{region 'Documentation'}
(*!
<summary>Selects explicit stimuli and expected results for one scenario.</summary>
*)
{endregion}
METHOD PRIVATE SelectScenario : BOOL //! TRUE after selecting a supported scenario and its literal expectations; FALSE reports an unknown scenario.
VAR
    Index : UINT;
END_VAR
SelectScenario := FALSE;
FSubjectEnable := TRUE;
FContinueScenario := FALSE;
FInput := 'A';
FExpected := 'B';
FWideInput := "A";
FWideExpected := "B";
FChar := BYTE#16#41;
FExpectedChar := BYTE#16#42;
FWideChar := WORD#16#0041;
FExpectedWideChar := WORD#16#0042;
CASE FScenario OF
    ScenarioShortQuoted:
        FExpectedMessage1 := 'Assertion failed: values are not equal. Expected = $'B$', Actual = $'A$'.';
        FExpectedMessage2 := 'Assertion failed: values are not equal. Expected = $'B$', Actual = $'A$'.';
        FExpectedMessage3 := 'Assertion failed: values are not equal. Expected = $'B$' (16#42), Actual = $'A$' (16#41).';
        FExpectedMessage4 := 'Assertion failed: values are not equal. Expected = $'B$' (16#0042), Actual = $'A$' (16#0041).';
        FTextExpectedResult := E_Result.Failed;
        FTextExpectedFinding := TRUE;
        FWideTextExpectedResult := E_Result.Failed;
        FWideTextExpectedFinding := TRUE;
        FCharacterExpectedResult := E_Result.Failed;
        FCharacterExpectedFinding := TRUE;
        FWideCharacterExpectedResult := E_Result.Failed;
        FWideCharacterExpectedFinding := TRUE;
    ScenarioPreview38:
        FInput := 'AAAAAAAAAAAAAAAAAAAAAAAAAAAAAAAAAAAAAA';
        FExpected := 'BBBBBBBBBBBBBBBBBBBBBBBBBBBBBBBBBBBBBB';
        FWideInput := "AAAAAAAAAAAAAAAAAAAAAAAAAAAAAAAAAAAAAA";
        FWideExpected := "BBBBBBBBBBBBBBBBBBBBBBBBBBBBBBBBBBBBBB";
        FExpectedMessage1 := 'Assertion failed: values are not equal. Expected = $'BBBBBBBBBBBBBBBBBBBBBBBBBBBBBBBBBBBBBB$', Actual = $'AAAAAAAAAAAAAAAAAAAAAAAAAAAAAAAAAAAAAA$'.';
        FExpectedMessage2 := 'Assertion failed: values are not equal. Expected = $'BBBBBBBBBBBBBBBBBBBBBBBBBBBBBBBBBBBBBB$', Actual = $'AAAAAAAAAAAAAAAAAAAAAAAAAAAAAAAAAAAAAA$'.';
        FExpectedMessage3 := 'Assertion failed: values are not equal. Expected = $'B$' (16#42), Actual = $'A$' (16#41).';
        FExpectedMessage4 := 'Assertion failed: values are not equal. Expected = $'B$' (16#0042), Actual = $'A$' (16#0041).';
        FTextExpectedResult := E_Result.Failed;
        FTextExpectedFinding := TRUE;
        FWideTextExpectedResult := E_Result.Failed;
        FWideTextExpectedFinding := TRUE;
        FCharacterExpectedResult := E_Result.Failed;
        FCharacterExpectedFinding := TRUE;
        FWideCharacterExpectedResult := E_Result.Failed;
        FWideCharacterExpectedFinding := TRUE;
    ScenarioPreview39:
        FInput := 'AAAAAAAAAAAAAAAAAAAAAAAAAAAAAAAAAAAAAAA';
        FExpected := 'BBBBBBBBBBBBBBBBBBBBBBBBBBBBBBBBBBBBBBB';
        FWideInput := "AAAAAAAAAAAAAAAAAAAAAAAAAAAAAAAAAAAAAAA";
        FWideExpected := "BBBBBBBBBBBBBBBBBBBBBBBBBBBBBBBBBBBBBBB";
        FExpectedMessage1 := 'Assertion failed: values are not equal. Expected = $'BBBBBBBBBBBBBBBBBBBBBBBBBBBBBBBBBBB...$', Actual = $'AAAAAAAAAAAAAAAAAAAAAAAAAAAAAAAAAAA...$'.';
        FExpectedMessage2 := 'Assertion failed: values are not equal. Expected = $'BBBBBBBBBBBBBBBBBBBBBBBBBBBBBBBBBBB...$', Actual = $'AAAAAAAAAAAAAAAAAAAAAAAAAAAAAAAAAAA...$'.';
        FExpectedMessage3 := 'Assertion failed: values are not equal. Expected = $'B$' (16#42), Actual = $'A$' (16#41).';
        FExpectedMessage4 := 'Assertion failed: values are not equal. Expected = $'B$' (16#0042), Actual = $'A$' (16#0041).';
        FTextExpectedResult := E_Result.Failed;
        FTextExpectedFinding := TRUE;
        FWideTextExpectedResult := E_Result.Failed;
        FWideTextExpectedFinding := TRUE;
        FCharacterExpectedResult := E_Result.Failed;
        FCharacterExpectedFinding := TRUE;
        FWideCharacterExpectedResult := E_Result.Failed;
        FWideCharacterExpectedFinding := TRUE;
    ScenarioDifferenceBeyondPreview:
        FInput := 'AAAAAAAAAAAAAAAAAAAAAAAAAAAAAAAAAAAAAAAX';
        FExpected := 'AAAAAAAAAAAAAAAAAAAAAAAAAAAAAAAAAAAAAAAY';
        FWideInput := "AAAAAAAAAAAAAAAAAAAAAAAAAAAAAAAAAAAAAAAX";
        FWideExpected := "AAAAAAAAAAAAAAAAAAAAAAAAAAAAAAAAAAAAAAAY";
        FExpectedMessage1 := 'Assertion failed: values are not equal. Expected = $'AAAAAAAAAAAAAAAAAAAAAAAAAAAAAAAAAAA...$', Actual = $'AAAAAAAAAAAAAAAAAAAAAAAAAAAAAAAAAAA...$'.';
        FExpectedMessage2 := 'Assertion failed: values are not equal. Expected = $'AAAAAAAAAAAAAAAAAAAAAAAAAAAAAAAAAAA...$', Actual = $'AAAAAAAAAAAAAAAAAAAAAAAAAAAAAAAAAAA...$'.';
        FExpectedMessage3 := 'Assertion failed: values are not equal. Expected = $'B$' (16#42), Actual = $'A$' (16#41).';
        FExpectedMessage4 := 'Assertion failed: values are not equal. Expected = $'B$' (16#0042), Actual = $'A$' (16#0041).';
        FTextExpectedResult := E_Result.Failed;
        FTextExpectedFinding := TRUE;
        FWideTextExpectedResult := E_Result.Failed;
        FWideTextExpectedFinding := TRUE;
        FCharacterExpectedResult := E_Result.Failed;
        FCharacterExpectedFinding := TRUE;
        FWideCharacterExpectedResult := E_Result.Failed;
        FWideCharacterExpectedFinding := TRUE;
    ScenarioAtCapacity:
        FOR Index := 0 TO Param_Assertions.AssertionStringLength - 1 DO
            // SA0175: Bounded byte writes construct exact input/terminator boundaries; no UTF-8 decoding.
            {analysis -175}
            FInput[Index] := BYTE#16#41;
            FExpected[Index] := BYTE#16#42;
            {analysis +175}
        END_FOR;
        // SA0175: Bounded byte writes construct exact input/terminator boundaries; no UTF-8 decoding.
        {analysis -175}
        FInput[Param_Assertions.AssertionStringLength] := 0;
        FExpected[Param_Assertions.AssertionStringLength] := 0;
        {analysis +175}
        FOR Index := 0 TO Param_Assertions.AssertionWStringLength - 1 DO
            FWideInput[Index] := WORD#16#0041;
            FWideExpected[Index] := WORD#16#0042;
        END_FOR;
        FWideInput[Param_Assertions.AssertionWStringLength] := 0;
        FWideExpected[Param_Assertions.AssertionWStringLength] := 0;
        FExpectedMessage1 := 'Assertion failed: values are not equal. Expected = $'BBBBBBBBBBBBBBBBBBBBBBBBBBBBBBBBBBB...$', Actual = $'AAAAAAAAAAAAAAAAAAAAAAAAAAAAAAAAAAA...$'.';
        FExpectedMessage2 := 'Assertion failed: values are not equal. Expected = $'BBBBBBBBBBBBBBBBBBBBBBBBBBBBBBBBBBB...$', Actual = $'AAAAAAAAAAAAAAAAAAAAAAAAAAAAAAAAAAA...$'.';
        FExpectedMessage3 := 'Assertion failed: values are not equal. Expected = $'B$' (16#42), Actual = $'A$' (16#41).';
        FExpectedMessage4 := 'Assertion failed: values are not equal. Expected = $'B$' (16#0042), Actual = $'A$' (16#0041).';
        FTextExpectedResult := E_Result.Failed;
        FTextExpectedFinding := TRUE;
        FWideTextExpectedResult := E_Result.Failed;
        FWideTextExpectedFinding := TRUE;
        FCharacterExpectedResult := E_Result.Failed;
        FCharacterExpectedFinding := TRUE;
        FWideCharacterExpectedResult := E_Result.Failed;
        FWideCharacterExpectedFinding := TRUE;
    ScenarioCodeFallback:
        FChar := 0;
        FExpectedChar := 1;
        FWideChar := WORD#16#0100;
        FExpectedWideChar := WORD#16#0200;
        FExpectedMessage1 := 'Assertion failed: values are not equal. Expected = $'B$', Actual = $'A$'.';
        FExpectedMessage2 := 'Assertion failed: values are not equal. Expected = $'B$', Actual = $'A$'.';
        FExpectedMessage3 := 'Assertion failed: values are not equal. Expected = 16#01, Actual = 16#00.';
        FExpectedMessage4 := 'Assertion failed: values are not equal. Expected = 16#0200, Actual = 16#0100.';
        FTextExpectedResult := E_Result.Failed;
        FTextExpectedFinding := TRUE;
        FWideTextExpectedResult := E_Result.Failed;
        FWideTextExpectedFinding := TRUE;
        FCharacterExpectedResult := E_Result.Failed;
        FCharacterExpectedFinding := TRUE;
        FWideCharacterExpectedResult := E_Result.Failed;
        FWideCharacterExpectedFinding := TRUE;
    ScenarioReplacement:
        // SA0175: Deliberately different raw bytes; both previews must render the same marker.
        {analysis -175}
        FInput := '$E4$01';
        FExpected := '$FF$7F';
        FWideInput := "$0100$20AC";
        FWideExpected := "$0001$FFFF";
        FExpectedMessage1 := 'Assertion failed: values are not equal. Expected = $'$D7$D7$', Actual = $'$D7$D7$'.';
        FExpectedMessage2 := 'Assertion failed: values are not equal. Expected = $'$D7$D7$', Actual = $'$D7$D7$'.';
        FExpectedMessage3 := 'Assertion failed: values are not equal. Expected = $'B$' (16#42), Actual = $'A$' (16#41).';
        FExpectedMessage4 := 'Assertion failed: values are not equal. Expected = $'B$' (16#0042), Actual = $'A$' (16#0041).';
        FTextExpectedResult := E_Result.Failed;
        FTextExpectedFinding := TRUE;
        FWideTextExpectedResult := E_Result.Failed;
        FWideTextExpectedFinding := TRUE;
        FCharacterExpectedResult := E_Result.Failed;
        FCharacterExpectedFinding := TRUE;
        FWideCharacterExpectedResult := E_Result.Failed;
        FWideCharacterExpectedFinding := TRUE;
        {analysis +175}
ELSE
    Error(Message := 'Unknown Assertion scenario.');
    RETURN;
END_CASE;
SelectScenario := TRUE;
END_METHOD

END_FUNCTION_BLOCK

// ---- Framework/Assertions/POU/Utilities/CreateAssertionTextValue_String.TcPOU
{region 'Documentation'}
(*!
<summary>Render a quoted diagnostic preview with at most AssertionValueLength output bytes.
Printable ASCII is retained; other code units become byte 16#D7 without expansion.</summary>
<description>
Zero terminates the input. Quotes and backslashes remain literal. Shortening reserves
space for enclosing quotes and an ellipsis; the default limit retains 35 code units.
Rendering is lossy and does not alter the compared input or its result.
</description>
*)
{endregion}
FUNCTION INTERNAL CreateAssertionTextValue_String : STRING(GVL_Constants.AssertionValueLength) //! Bounded diagnostic aid; not a lossless representation for subsequent comparison.
VAR_INPUT
    Value : STRING(GVL_Constants.MessageLength); //! Text to preview; zero terminates the input.
END_VAR
VAR
    Text : STRING(GVL_Constants.AssertionValueLength);
    CharacterIndex : INT;
    CopyLength : INT;
    Code : BYTE;
    Shortened : BOOL;
END_VAR
VAR CONSTANT
    Quote : STRING(1) := '$'';
    Ellipsis : STRING(3) := '...';
    QuoteLength : INT := 2;
    EllipsisLength : INT := 3;
    FirstPrintableAscii : BYTE := 16#20;
    LastPrintableAscii : BYTE := 16#7E;
    ReplacementByte : BYTE := 16#D7;
END_VAR

CopyLength := UINT_TO_INT(GVL_Constants.AssertionValueLength) - QuoteLength;
// SA0175: Bounded diagnostic code-unit rendering; each unsupported unit becomes one byte.
{analysis -175}
Shortened := TRUE;
FOR CharacterIndex := 0 TO CopyLength DO
    IF Value[CharacterIndex] = 0 THEN
        CopyLength := CharacterIndex;
        Shortened := FALSE;
        EXIT;
    END_IF;
END_FOR;
IF Shortened THEN
    CopyLength := CopyLength - EllipsisLength;
END_IF;

FOR CharacterIndex := 0 TO CopyLength - 1 DO
    Code := Value[CharacterIndex];
    IF (Code >= FirstPrintableAscii) AND (Code <= LastPrintableAscii) THEN
        Text[CharacterIndex] := Code;
    ELSE
        Text[CharacterIndex] := ReplacementByte;
    END_IF;
END_FOR;
Text[CopyLength] := 0;
{analysis +175}

IF Shortened THEN
    Text := CONCAT(Text, Ellipsis);
END_IF;
CreateAssertionTextValue_String := CONCAT(Quote, Text);
CreateAssertionTextValue_String := CONCAT(CreateAssertionTextValue_String, Quote);

END_FUNCTION

// ---- Framework/Assertions/POU/Utilities/CreateAssertionTextValue_WString.TcPOU
{region 'Documentation'}
(*!
<summary>Render a quoted diagnostic preview with at most AssertionValueLength output bytes.
Printable ASCII is retained; other code units become byte 16#D7 without expansion.</summary>
<description>
Zero terminates the input. Quotes and backslashes remain literal. Shortening reserves
space for enclosing quotes and an ellipsis; the default limit retains 35 code units.
Rendering is lossy and does not alter the compared input or its result.
</description>
*)
{endregion}
FUNCTION INTERNAL CreateAssertionTextValue_WString : STRING(GVL_Constants.AssertionValueLength) //! Bounded diagnostic aid; not a lossless representation for subsequent comparison.
VAR_INPUT
    Value : WSTRING(GVL_Constants.MessageLength); //! Text to preview; zero terminates the input.
END_VAR
VAR
    Text : STRING(GVL_Constants.AssertionValueLength);
    CharacterIndex : INT;
    CopyLength : INT;
    Code : WORD;
    Shortened : BOOL;
END_VAR
VAR CONSTANT
    Quote : STRING(1) := '$'';
    Ellipsis : STRING(3) := '...';
    QuoteLength : INT := 2;
    EllipsisLength : INT := 3;
    FirstPrintableAscii : WORD := 16#20;
    LastPrintableAscii : WORD := 16#7E;
    ReplacementByte : BYTE := 16#D7;
END_VAR

CopyLength := UINT_TO_INT(GVL_Constants.AssertionValueLength) - QuoteLength;
// SA0175: Bounded diagnostic code-unit rendering; each unsupported unit becomes one byte.
{analysis -175}
Shortened := TRUE;
FOR CharacterIndex := 0 TO CopyLength DO
    IF Value[CharacterIndex] = 0 THEN
        CopyLength := CharacterIndex;
        Shortened := FALSE;
        EXIT;
    END_IF;
END_FOR;
IF Shortened THEN
    CopyLength := CopyLength - EllipsisLength;
END_IF;

FOR CharacterIndex := 0 TO CopyLength - 1 DO
    Code := Value[CharacterIndex];
    IF (Code >= FirstPrintableAscii) AND (Code <= LastPrintableAscii) THEN
        Text[CharacterIndex] := WORD_TO_BYTE(Code);
    ELSE
        Text[CharacterIndex] := ReplacementByte;
    END_IF;
END_FOR;
Text[CopyLength] := 0;
{analysis +175}

IF Shortened THEN
    Text := CONCAT(Text, Ellipsis);
END_IF;
CreateAssertionTextValue_WString := CONCAT(Quote, Text);
CreateAssertionTextValue_WString := CONCAT(CreateAssertionTextValue_WString, Quote);

END_FUNCTION

// ---- Framework/Assertions/POU/Utilities/CreateAssertionTextValue_ByteArray.TcPOU
{region 'Documentation'}
(*!
<summary>Render a quoted printable-ASCII/16#D7 preview of an array range without modifying its storage. Invalid or empty ranges return two quotes. Zero and other unsupported elements become one replacement byte each. Work is bounded by the preview capacity.</summary>
*)
{endregion}
FUNCTION INTERNAL CreateAssertionTextValue_ByteArray : STRING(GVL_Constants.AssertionValueLength) //! Bounded diagnostic text; not a value for subsequent numeric comparison.
VAR_INPUT
    StartIndex : DINT; //! First selected index in Value, using the array's declared index range.
    Length : UINT; //! Number of selected elements starting at StartIndex; must fit the array range.
END_VAR
VAR_IN_OUT CONSTANT
    Value : ARRAY[*] OF BYTE; //! Read-only source array; StartIndex and Length select the diagnostic preview.
END_VAR
VAR
    LowerIndex : DINT;
    UpperIndex : DINT;
    CopyLength : INT;
    Offset : INT;
    Code : BYTE;
    Text : STRING(GVL_Constants.AssertionValueLength);
    Preview : STRING(GVL_Constants.AssertionValueLength);
END_VAR
VAR CONSTANT
    Quote : STRING(1) := '$'';
    Ellipsis : STRING(3) := '...';
    QuoteLength : INT := 2;
    EllipsisLength : INT := 3;
    FirstPrintableAscii : BYTE := 16#20;
    LastPrintableAscii : BYTE := 16#7E;
    ReplacementByte : BYTE := 16#D7;
END_VAR

CreateAssertionTextValue_ByteArray := CONCAT(Quote, Quote);
LowerIndex := LOWER_BOUND(Value, 1);
UpperIndex := UPPER_BOUND(Value, 1);

IF Length = 0 OR StartIndex < LowerIndex OR StartIndex > UpperIndex THEN
    RETURN;
END_IF;

IF UINT_TO_LINT(Length) > DINT_TO_LINT(UpperIndex) - DINT_TO_LINT(StartIndex) + 1 THEN
    RETURN;
END_IF;

IF Length > GVL_Constants.AssertionValueLength - INT_TO_UINT(QuoteLength) THEN
    CopyLength := UINT_TO_INT(GVL_Constants.AssertionValueLength) - QuoteLength - EllipsisLength;
ELSE
    CopyLength := UINT_TO_INT(Length);
END_IF;

// SA0175: Range guards bound reads; preview writes fit capacity, including the terminator.
{analysis -175}
FOR Offset := 0 TO CopyLength - 1 DO
    Code := Value[StartIndex + INT_TO_DINT(Offset)];
    IF (Code >= FirstPrintableAscii) AND (Code <= LastPrintableAscii) THEN
        Text[Offset] := Code;
    ELSE
        Text[Offset] := ReplacementByte;
    END_IF;
END_FOR;
Text[CopyLength] := 0;
{analysis +175}

Preview := Text;
IF Length > GVL_Constants.AssertionValueLength - INT_TO_UINT(QuoteLength) THEN
    Preview := CONCAT(Preview, Ellipsis);
END_IF;

CreateAssertionTextValue_ByteArray := CONCAT(Quote, Preview);
CreateAssertionTextValue_ByteArray := CONCAT(CreateAssertionTextValue_ByteArray, Quote);

END_FUNCTION

// ---- Framework/Assertions/POU/Utilities/CreateAssertionTextValue_WordArray.TcPOU
{region 'Documentation'}
(*!
<summary>Render a quoted printable-ASCII/16#D7 preview of an array range without modifying its storage. Invalid or empty ranges return two quotes. Zero and other unsupported elements become one replacement byte each. Work is bounded by the preview capacity.</summary>
*)
{endregion}
FUNCTION INTERNAL CreateAssertionTextValue_WordArray : STRING(GVL_Constants.AssertionValueLength) //! Bounded diagnostic text; not a value for subsequent numeric comparison.
VAR_INPUT
    StartIndex : DINT; //! First selected index in Value, using the array's declared index range.
    Length : UINT; //! Number of selected elements starting at StartIndex; must fit the array range.
END_VAR
VAR_IN_OUT CONSTANT
    Value : ARRAY[*] OF WORD; //! Read-only source array; StartIndex and Length select the diagnostic preview.
END_VAR
VAR
    LowerIndex : DINT;
    UpperIndex : DINT;
    CopyLength : INT;
    Offset : INT;
    Code : WORD;
    Text : STRING(GVL_Constants.AssertionValueLength);
    Preview : STRING(GVL_Constants.AssertionValueLength);
END_VAR
VAR CONSTANT
    Quote : STRING(1) := '$'';
    Ellipsis : STRING(3) := '...';
    QuoteLength : INT := 2;
    EllipsisLength : INT := 3;
    FirstPrintableAscii : WORD := 16#20;
    LastPrintableAscii : WORD := 16#7E;
    ReplacementByte : BYTE := 16#D7;
END_VAR

CreateAssertionTextValue_WordArray := CONCAT(Quote, Quote);
LowerIndex := LOWER_BOUND(Value, 1);
UpperIndex := UPPER_BOUND(Value, 1);

IF Length = 0 OR StartIndex < LowerIndex OR StartIndex > UpperIndex THEN
    RETURN;
END_IF;

IF UINT_TO_LINT(Length) > DINT_TO_LINT(UpperIndex) - DINT_TO_LINT(StartIndex) + 1 THEN
    RETURN;
END_IF;

IF Length > GVL_Constants.AssertionValueLength - INT_TO_UINT(QuoteLength) THEN
    CopyLength := UINT_TO_INT(GVL_Constants.AssertionValueLength) - QuoteLength - EllipsisLength;
ELSE
    CopyLength := UINT_TO_INT(Length);
END_IF;

// SA0175: Range guards bound reads; preview writes fit capacity, including the terminator.
{analysis -175}
FOR Offset := 0 TO CopyLength - 1 DO
    Code := Value[StartIndex + INT_TO_DINT(Offset)];
    IF (Code >= FirstPrintableAscii) AND (Code <= LastPrintableAscii) THEN
        Text[Offset] := WORD_TO_BYTE(Code);
    ELSE
        Text[Offset] := ReplacementByte;
    END_IF;
END_FOR;
Text[CopyLength] := 0;
{analysis +175}

Preview := Text;
IF Length > GVL_Constants.AssertionValueLength - INT_TO_UINT(QuoteLength) THEN
    Preview := CONCAT(Preview, Ellipsis);
END_IF;

CreateAssertionTextValue_WordArray := CONCAT(Quote, Preview);
CreateAssertionTextValue_WordArray := CONCAT(CreateAssertionTextValue_WordArray, Quote);

END_FUNCTION

// ---- Framework/Assertions/POU/Utilities/CreateAssertionTextValue_WChar.TcPOU
{region 'Documentation'}
(*!
<summary>Formats printable ASCII as a quoted character and hexadecimal code; other values as code only. Output is ASCII and at most 13 characters.</summary>
*)
{endregion}
FUNCTION INTERNAL CreateAssertionTextValue_WChar : STRING(13) //! Bounded diagnostic text; not a value for subsequent numeric comparison.
VAR_INPUT
    Value : WORD; //! Character code to render; no character validation is performed.
END_VAR
VAR
    HexText : STRING(7);
    Text : STRING(13);
END_VAR
VAR CONSTANT
    FirstPrintableAscii : WORD := 16#20;
    LastPrintableAscii : WORD := 16#7E;
    HexDigitCount : USINT := 4;
END_VAR

HexText := CreateAssertionTextValue_Hex(Value := WORD_TO_LWORD(Value),
    DigitCount := HexDigitCount);

IF (Value < FirstPrintableAscii) OR (Value > LastPrintableAscii) THEN
    CreateAssertionTextValue_WChar := HexText;
    RETURN;
END_IF;

Text := '$' $' (';
// SA0175: Printable-ASCII guard; index 1 fits the quoted template.
{analysis -175}
Text[1] := WORD_TO_BYTE(Value);
{analysis +175}
Text := CONCAT(Text, HexText);
CreateAssertionTextValue_WChar := CONCAT(Text, ')');

END_FUNCTION

// ---- SelfTests/TestCases/TestSuite_AssertionText/Test_AssertionValueTokenCount.TcPOU
{region 'Documentation'}
(*!
<summary>Checks masked BYTE/WORD token counts, count predicates and retained observations.</summary>
<description>
Literal counts distinguish full masks, selected bits, zero mask and sliced ranges.
Dedicated continuation scenarios check disabled/Failed count retention and clearing
on invalid range. Every independent scenario verifies count clearing on Reset.
Independent scenarios occupy two calls: bound Reset, then evaluation.
ProcessAssertions checks each call before ProcessTests advances. Literal expected
results belong to SelectScenario, not to a copy of the production comparison.
The local capture is cleared before each call and checked in subject-call order.
FirstFailedScenario and FailedDuringEvaluation retain the first mismatch.
Continuation scenarios explicitly retain the prior subject state. The Test Case
owns all input storage; no invalid or dangling references are constructed.
</description>
*)
{endregion}
FUNCTION_BLOCK Test_AssertionValueTokenCount EXTENDS TestCaseBase
VAR
    FEqual : AssertValueTokenCntEqual_Byte;
    FEqualExpectedResult : E_Result;
    FWideEqual : AssertValueTokenCntEqual_Word;
    FWideEqualExpectedResult : E_Result;
    FNone : AssertNoValueToken_Byte;
    FNoneExpectedResult : E_Result;
    FWideRange : AssertValueTokenCntInRange_Word;
    FWideRangeExpectedResult : E_Result;
    FData : ARRAY[-2..3] OF BYTE;
    FDataBefore : ARRAY[-2..3] OF BYTE;
    FWideData : ARRAY[-2..3] OF WORD;
    FWideDataBefore : ARRAY[-2..3] OF WORD;
    FStartIndex : DINT;
    FLength : USINT;
    FExpected : UINT;
    FMinimum : UINT;
    FMaximum : UINT;
    FToken : BYTE;
    FWideToken : WORD;
    FMask : BYTE;
    FWideMask : WORD;
    FSubjectEnable : BOOL;
    FContinueScenario : BOOL;
    FEqualExpectedFinding : BOOL;
    FEqualExpectedCount : UINT;
    FWideEqualExpectedFinding : BOOL;
    FWideEqualExpectedCount : UINT;
    FNoneExpectedFinding : BOOL;
    FNoneExpectedCount : UINT;
    FWideRangeExpectedFinding : BOOL;
    FWideRangeExpectedCount : UINT;
    FCapture : EventBuffer;
    FEvents : ARRAY[1..CaptureLength] OF ST_Event;
    FCaptureFifo : ST_FifoStatus;
    FCaptureStatus : ST_EventBufferStatus;
    FSetupValid : BOOL;
    FScenario : UINT;
    FChecked : BOOL;
    FEvaluateSubjects : BOOL;
    FObservationReady : BOOL;
    FFirstFailedScenario : UINT;
    FFailedDuringEvaluation : BOOL;
    FResultsMatch : BOOL;
    FResults : AssertTrue;
    FActivityMatch : BOOL;
    FActivity : AssertTrue;
    FInputsMatch : BOOL;
    FInputs : AssertTrue;
    FFindingsMatch : BOOL;
    FFindings : AssertTrue;
END_VAR
VAR CONSTANT
    CaptureLength : UINT := 8;
    ScenarioExactCount : UINT := 1;
    ScenarioMasked : UINT := 2;
    ScenarioZeroMask : UINT := 3;
    ScenarioSelectedBounds : UINT := 4;
    ScenarioLastElement : UINT := 5;
    ScenarioAbsent : UINT := 6;
    ScenarioFailedCount : UINT := 7;
    ScenarioDisabledRetention : UINT := 8;
    ScenarioFailedRetention : UINT := 9;
    ScenarioErrorClearsCount : UINT := 10;
    ScenarioResetAfterError : UINT := 11;
    ScenarioBelowArray : UINT := 12;
    ScenarioEndOutsideArray : UINT := 13;
    ScenarioReversedCountBounds : UINT := 14;
    LastScenario : UINT := ScenarioReversedCountBounds;
END_VAR

SUPER^();

{region 'Documentation'}
(*!
<summary>Aggregates only outer checks, not intentionally failing subjects.</summary>
*)
{endregion}
METHOD PROTECTED AggregateResults
VAR_INPUT
    Aggregator : I_ResultAggregator; //! Borrowed result sink owned by the outer Test Case; add this test's checking Assertions without resetting or retaining the sink.
END_VAR
Aggregator.AddProvider(Provider := FResults);
Aggregator.AddProvider(Provider := FActivity);
Aggregator.AddProvider(Provider := FInputs);
Aggregator.AddProvider(Provider := FFindings);
END_METHOD

{region 'Documentation'}
(*!
<summary>Calls each inherited production subject once with caller-owned input storage.</summary>
*)
{endregion}
METHOD PRIVATE CallSubjects
FEqual(Enable := FSubjectEnable,
    State := E_State.Running,
    StartIndex := FStartIndex,
    Length := FLength,
    Expected := FExpected,
    Token := FToken,
    Mask := FMask,
    IN := FData);
FWideEqual(Enable := FSubjectEnable,
    State := E_State.Running,
    StartIndex := FStartIndex,
    Length := FLength,
    Expected := FExpected,
    Token := FWideToken,
    Mask := FWideMask,
    IN := FWideData);
FNone(Enable := FSubjectEnable,
    State := E_State.Running,
    StartIndex := FStartIndex,
    Length := FLength,
    Token := FToken,
    Mask := FMask,
    IN := FData);
FWideRange(Enable := FSubjectEnable,
    State := E_State.Running,
    StartIndex := FStartIndex,
    Length := FLength,
    Minimum := FMinimum,
    Maximum := FMaximum,
    Token := FWideToken,
    Mask := FWideMask,
    IN := FWideData);
END_METHOD

{region 'Documentation'}
(*!
<summary>Checks one subject finding in call order; expected outcomes come from the scenario.</summary>
*)
{endregion}
METHOD PRIVATE CheckFinding : BOOL //! TRUE when the required finding checks pass; calls requiring no finding also succeed.
VAR_INPUT
    Subject : I_Assertion; //! Assertion interface supplying the expected finding identity.
    ExpectedResult : E_Result; //! Independently authored result expected in the captured finding.
    ExpectedFinding : BOOL; //! TRUE when this scenario requires a finding during active evaluation.
END_VAR
VAR_IN_OUT
    Index : UINT; //! One-based next finding index; advanced when this call checks a required finding.
END_VAR
CheckFinding := TRUE;
IF FEvaluateSubjects AND ExpectedFinding THEN
    CheckFinding := (FEvents[Index].SequenceId = UINT_TO_UDINT(Index))
        AND (FEvents[Index].Name = Subject.Name)
        AND (FEvents[Index].OwnerScope = E_OwnerScope.Assertion)
        AND (FEvents[Index].EventType = E_EventType.Result)
        AND (FEvents[Index].State = E_State.Running)
        AND (FEvents[Index].Result = ExpectedResult)
        AND (FEvents[Index].Message <> '');
    Index := Index + 1;
END_IF;
END_METHOD

{region 'Documentation'}
(*!
<summary>Checks exact finding count and identities; at most one finding per subject.</summary>
*)
{endregion}
METHOD PRIVATE CheckFindings
VAR
    Index : UINT;
    Matches : BOOL;
END_VAR
Index := 1;
FFindingsMatch := TRUE;
Matches := CheckFinding(Subject := FEqual,
    ExpectedResult := FEqualExpectedResult,
    ExpectedFinding := FEqualExpectedFinding,
    Index := Index);
FFindingsMatch := FFindingsMatch AND Matches;
Matches := CheckFinding(Subject := FWideEqual,
    ExpectedResult := FWideEqualExpectedResult,
    ExpectedFinding := FWideEqualExpectedFinding,
    Index := Index);
FFindingsMatch := FFindingsMatch AND Matches;
Matches := CheckFinding(Subject := FNone,
    ExpectedResult := FNoneExpectedResult,
    ExpectedFinding := FNoneExpectedFinding,
    Index := Index);
FFindingsMatch := FFindingsMatch AND Matches;
Matches := CheckFinding(Subject := FWideRange,
    ExpectedResult := FWideRangeExpectedResult,
    ExpectedFinding := FWideRangeExpectedFinding,
    Index := Index);
FFindingsMatch := FFindingsMatch AND Matches;
FFindingsMatch := FFindingsMatch
    AND (FCaptureStatus.SequenceId = UINT_TO_UDINT(Index - 1))
    AND (FCaptureStatus.LostEventCount = 0);
IF FEvaluateSubjects AND (FScenario = ScenarioFailedCount) THEN
    // SA0175: Fixed byte-substring checks of bounded diagnostic messages; no character offsets.
    {analysis -175}
    FFindingsMatch := FFindingsMatch
        AND (FIND(FEvents[1].Message, 'Actual = 2') > 0)
        AND (FIND(FEvents[4].Message, 'Actual = 2') > 0);
    {analysis +175}
END_IF;
END_METHOD

{region 'Documentation'}
(*!
<summary>Rejects incomplete subject, capture or outer Assertion setup.</summary>
*)
{endregion}
METHOD PROTECTED CheckInitialization : BOOL //! TRUE when the inherited initialization check and this concrete fixture check both accept the setup.
CheckInitialization := SUPER^.CheckInitialization();
IF NOT CheckInitialization THEN
    RETURN;
END_IF;

CheckInitialization := FSetupValid
    AND FResults.IsInitialized
    AND FActivity.IsInitialized
    AND FInputs.IsInitialized
    AND FFindings.IsInitialized;
IF NOT CheckInitialization THEN
    EventPublisher.PublishEvent(Event := CreateFrameworkEvent(Name := Name,
        ResourceName := '',
        State := State,
        Severity := E_EventSeverity.Error,
        Message := 'Text selftest setup failed.'));
END_IF;
END_METHOD

{region 'Documentation'}
(*!
<summary>Checks literal evaluation results, or NotEvaluated on the reset call.</summary>
*)
{endregion}
METHOD PRIVATE CheckResults
IF FEvaluateSubjects THEN
    FResultsMatch := (FEqual.Result = FEqualExpectedResult)
        AND (FWideEqual.Result = FWideEqualExpectedResult)
        AND (FNone.Result = FNoneExpectedResult)
        AND (FWideRange.Result = FWideRangeExpectedResult);
ELSE
    FResultsMatch := (FEqual.Result = E_Result.NotEvaluated)
        AND (FWideEqual.Result = E_Result.NotEvaluated)
        AND (FNone.Result = E_Result.NotEvaluated)
        AND (FWideRange.Result = E_Result.NotEvaluated);
END_IF;
FActivityMatch := (FEqual.Enabled = FSubjectEnable)
    AND (FEqual.ObservationActive = (FEvaluateSubjects AND FSubjectEnable))
    AND (FEqual.EvaluationActive = (FEvaluateSubjects AND FSubjectEnable))
    AND (FWideEqual.Enabled = FSubjectEnable)
    AND (FWideEqual.ObservationActive = (FEvaluateSubjects AND FSubjectEnable))
    AND (FWideEqual.EvaluationActive = (FEvaluateSubjects AND FSubjectEnable))
    AND (FNone.Enabled = FSubjectEnable)
    AND (FNone.ObservationActive = (FEvaluateSubjects AND FSubjectEnable))
    AND (FNone.EvaluationActive = (FEvaluateSubjects AND FSubjectEnable))
    AND (FWideRange.Enabled = FSubjectEnable)
    AND (FWideRange.ObservationActive = (FEvaluateSubjects AND FSubjectEnable))
    AND (FWideRange.EvaluationActive = (FEvaluateSubjects AND FSubjectEnable));
IF FEvaluateSubjects THEN
    FResultsMatch := FResultsMatch
        AND (FEqual.TokenCount = FEqualExpectedCount)
        AND (FWideEqual.TokenCount = FWideEqualExpectedCount)
        AND (FNone.TokenCount = FNoneExpectedCount)
        AND (FWideRange.TokenCount = FWideRangeExpectedCount);
ELSE
    FResultsMatch := FResultsMatch
        AND (FEqual.TokenCount = 0)
        AND (FWideEqual.TokenCount = 0)
        AND (FNone.TokenCount = 0)
        AND (FWideRange.TokenCount = 0);
END_IF;
END_METHOD

{region 'Documentation'}
(*!
<summary>Initializes outer checks and isolates intentional subject findings.</summary>
*)
{endregion}
METHOD PROTECTED Configure
VAR
    Initialized : BOOL;
END_VAR
FPreparationStateCount := 0;
FTestStateCount := 1;
FResults.Initialize(Parent := THIS^,
    AssertionName := 'Results');
FActivity.Initialize(Parent := THIS^,
    AssertionName := 'Activity');
FInputs.Initialize(Parent := THIS^,
    AssertionName := 'Inputs');
FFindings.Initialize(Parent := THIS^,
    AssertionName := 'Findings');
FSetupValid := FCapture.Initialize(Buffer := FEvents,
    FifoControl := FCaptureFifo,
    Status := FCaptureStatus);
FEqual.BindPublisher(Publisher := FCapture);
Initialized := FEqual.Initialize(Parent := THIS^,
    AssertionName := 'Equal');
FSetupValid := FSetupValid AND Initialized;
FWideEqual.BindPublisher(Publisher := FCapture);
Initialized := FWideEqual.Initialize(Parent := THIS^,
    AssertionName := 'WideEqual');
FSetupValid := FSetupValid AND Initialized;
FNone.BindPublisher(Publisher := FCapture);
Initialized := FNone.Initialize(Parent := THIS^,
    AssertionName := 'None');
FSetupValid := FSetupValid AND Initialized;
FWideRange.BindPublisher(Publisher := FCapture);
Initialized := FWideRange.Initialize(Parent := THIS^,
    AssertionName := 'WideRange');
FSetupValid := FSetupValid AND Initialized;
END_METHOD

{region 'Documentation'}
(*!
<summary>Completes abort; no asynchronous resource is owned.</summary>
*)
{endregion}
METHOD PROTECTED ProcessAbort
VAR_INPUT
    Enable : BOOL; //! Phase permission supplied by the owning Test Case; FALSE does not authorize progression, while observation may continue.
END_VAR
IF Enable THEN
    CompleteAbort();
END_IF;
END_METHOD

{region 'Documentation'}
(*!
<summary>Latches this call's checks before progression is permitted.</summary>
*)
{endregion}
METHOD PROTECTED ProcessAssertions
VAR_INPUT
    Enable : BOOL; //! Phase permission supplied by the owning Test Case; FALSE does not authorize progression, while observation may continue.
END_VAR
VAR
    Check : BOOL;
END_VAR
Check := Enable AND FObservationReady;
FResults(Enable := Check,
    State := State,
    IN := FResultsMatch);
FActivity(Enable := Check,
    State := State,
    IN := FActivityMatch);
FInputs(Enable := Check,
    State := State,
    IN := FInputsMatch);
FFindings(Enable := Check,
    State := State,
    IN := FFindingsMatch);
IF Check THEN
    FChecked := TRUE;
END_IF;
END_METHOD

{region 'Documentation'}
(*!
<summary>No Preparation phase is needed.</summary>
*)
{endregion}
METHOD PROTECTED ProcessPreparations
VAR_INPUT
    // SA0033: Required hook; this test has no Preparation phase.
    {attribute 'analysis' := '-33'}
    Enable : BOOL; //! Phase permission supplied by the owning Test Case; FALSE does not authorize progression, while observation may continue.
END_VAR
END_METHOD

{region 'Documentation'}
(*!
<summary>Restarts the scenario sequence and outer checks.</summary>
*)
{endregion}
METHOD PROTECTED ProcessReset
FScenario := ScenarioExactCount;
FChecked := FALSE;
FSubjectEnable := FALSE;
FContinueScenario := FALSE;
FEvaluateSubjects := FALSE;
FObservationReady := FALSE;
FFirstFailedScenario := 0;
FFailedDuringEvaluation := FALSE;
FCapture.Reset();
ResetSubjects();
FResults.Reset();
FActivity.Reset();
FInputs.Reset();
FFindings.Reset();
CompleteReset();
END_METHOD

{region 'Documentation'}
(*!
<summary>Consumes reset before each independent scenario; continuation retains subject state.</summary>
*)
{endregion}
METHOD PROTECTED ProcessTests
VAR_INPUT
    Enable : BOOL; //! Phase permission supplied by the owning Test Case; FALSE does not authorize progression, while observation may continue.
END_VAR
IF NOT Enable THEN
    RETURN;
END_IF;

IF FChecked THEN
    FChecked := FALSE;
    FObservationReady := FALSE;
    IF FEvaluateSubjects THEN
        IF FScenario = LastScenario THEN
            CompleteTests();
            RETURN;
        END_IF;
        FScenario := FScenario + 1;
    END_IF;
    FEvaluateSubjects := NOT FEvaluateSubjects;
END_IF;

IF NOT SelectScenario() THEN
    RETURN;
END_IF;
IF FContinueScenario THEN
    FEvaluateSubjects := TRUE;
END_IF;
FCapture.Reset();
IF NOT FEvaluateSubjects THEN
    ResetSubjects();
END_IF;
FDataBefore := FData;
FWideDataBefore := FWideData;
CallSubjects();
CheckResults();
FInputsMatch := (FData[-2] = FDataBefore[-2])
    AND (FData[-1] = FDataBefore[-1])
    AND (FData[0] = FDataBefore[0])
    AND (FData[1] = FDataBefore[1])
    AND (FData[2] = FDataBefore[2])
    AND (FData[3] = FDataBefore[3])
    AND (FWideData[-2] = FWideDataBefore[-2])
    AND (FWideData[-1] = FWideDataBefore[-1])
    AND (FWideData[0] = FWideDataBefore[0])
    AND (FWideData[1] = FWideDataBefore[1])
    AND (FWideData[2] = FWideDataBefore[2])
    AND (FWideData[3] = FWideDataBefore[3]);
CheckFindings();
IF (FFirstFailedScenario = 0)
    AND NOT (FResultsMatch AND FActivityMatch AND FInputsMatch AND FFindingsMatch) THEN
    FFirstFailedScenario := FScenario;
    FFailedDuringEvaluation := FEvaluateSubjects;
END_IF;
FObservationReady := TRUE;
END_METHOD

{region 'Documentation'}
(*!
<summary>Queues reset; the next bound FB call consumes it without evaluating.</summary>
*)
{endregion}
METHOD PRIVATE ResetSubjects
FEqual.Reset();
FWideEqual.Reset();
FNone.Reset();
FWideRange.Reset();
END_METHOD

{region 'Documentation'}
(*!
<summary>Selects explicit stimuli and expected results for one scenario.</summary>
*)
{endregion}
METHOD PRIVATE SelectScenario : BOOL //! TRUE after selecting a supported scenario and its literal expectations; FALSE reports an unknown scenario.
SelectScenario := FALSE;
FSubjectEnable := TRUE;
FContinueScenario := FALSE;
FData[-2] := BYTE#16#10;
FData[-1] := BYTE#16#21;
FData[0] := BYTE#16#11;
FData[1] := BYTE#16#20;
FData[2] := BYTE#16#11;
FData[3] := BYTE#16#99;
FWideData[-2] := WORD#16#0110;
FWideData[-1] := WORD#16#0121;
FWideData[0] := WORD#16#0111;
FWideData[1] := WORD#16#0220;
FWideData[2] := WORD#16#0111;
FWideData[3] := WORD#16#0099;
FStartIndex := -2;
FLength := 6;
FExpected := 2;
FMinimum := 2;
FMaximum := 2;
FToken := BYTE#16#11;
FWideToken := WORD#16#0111;
FMask := BYTE#16#FF;
FWideMask := WORD#16#FFFF;
CASE FScenario OF
    ScenarioExactCount:
        FEqualExpectedResult := E_Result.Passed;
        FEqualExpectedFinding := FALSE;
        FEqualExpectedCount := 2;
        FWideEqualExpectedResult := E_Result.Passed;
        FWideEqualExpectedFinding := FALSE;
        FWideEqualExpectedCount := 2;
        FNoneExpectedResult := E_Result.Failed;
        FNoneExpectedFinding := TRUE;
        FNoneExpectedCount := 2;
        FWideRangeExpectedResult := E_Result.Passed;
        FWideRangeExpectedFinding := FALSE;
        FWideRangeExpectedCount := 2;
    ScenarioMasked:
        FMask := BYTE#16#0F;
        FWideMask := WORD#16#000F;
        FExpected := 3;
        FMinimum := 3;
        FMaximum := 3;
        FEqualExpectedResult := E_Result.Passed;
        FEqualExpectedFinding := FALSE;
        FEqualExpectedCount := 3;
        FWideEqualExpectedResult := E_Result.Passed;
        FWideEqualExpectedFinding := FALSE;
        FWideEqualExpectedCount := 3;
        FNoneExpectedResult := E_Result.Failed;
        FNoneExpectedFinding := TRUE;
        FNoneExpectedCount := 3;
        FWideRangeExpectedResult := E_Result.Passed;
        FWideRangeExpectedFinding := FALSE;
        FWideRangeExpectedCount := 3;
    ScenarioZeroMask:
        FMask := 0;
        FWideMask := 0;
        FExpected := 6;
        FMinimum := 6;
        FMaximum := 6;
        FEqualExpectedResult := E_Result.Passed;
        FEqualExpectedFinding := FALSE;
        FEqualExpectedCount := 6;
        FWideEqualExpectedResult := E_Result.Passed;
        FWideEqualExpectedFinding := FALSE;
        FWideEqualExpectedCount := 6;
        FNoneExpectedResult := E_Result.Failed;
        FNoneExpectedFinding := TRUE;
        FNoneExpectedCount := 6;
        FWideRangeExpectedResult := E_Result.Passed;
        FWideRangeExpectedFinding := FALSE;
        FWideRangeExpectedCount := 6;
    ScenarioSelectedBounds:
        FStartIndex := 0;
        FLength := 3;
        FData[-2] := FToken;
        FData[3] := FToken;
        FWideData[-2] := FWideToken;
        FWideData[3] := FWideToken;
        FEqualExpectedResult := E_Result.Passed;
        FEqualExpectedFinding := FALSE;
        FEqualExpectedCount := 2;
        FWideEqualExpectedResult := E_Result.Passed;
        FWideEqualExpectedFinding := FALSE;
        FWideEqualExpectedCount := 2;
        FNoneExpectedResult := E_Result.Failed;
        FNoneExpectedFinding := TRUE;
        FNoneExpectedCount := 2;
        FWideRangeExpectedResult := E_Result.Passed;
        FWideRangeExpectedFinding := FALSE;
        FWideRangeExpectedCount := 2;
    ScenarioLastElement:
        FStartIndex := 3;
        FLength := 1;
        FToken := BYTE#16#99;
        FWideToken := WORD#16#0099;
        FExpected := 1;
        FMinimum := 1;
        FMaximum := 1;
        FEqualExpectedResult := E_Result.Passed;
        FEqualExpectedFinding := FALSE;
        FEqualExpectedCount := 1;
        FWideEqualExpectedResult := E_Result.Passed;
        FWideEqualExpectedFinding := FALSE;
        FWideEqualExpectedCount := 1;
        FNoneExpectedResult := E_Result.Failed;
        FNoneExpectedFinding := TRUE;
        FNoneExpectedCount := 1;
        FWideRangeExpectedResult := E_Result.Passed;
        FWideRangeExpectedFinding := FALSE;
        FWideRangeExpectedCount := 1;
    ScenarioAbsent:
        FToken := 0;
        FWideToken := 0;
        FExpected := 0;
        FMinimum := 0;
        FMaximum := 0;
        FEqualExpectedResult := E_Result.Passed;
        FEqualExpectedFinding := FALSE;
        FEqualExpectedCount := 0;
        FWideEqualExpectedResult := E_Result.Passed;
        FWideEqualExpectedFinding := FALSE;
        FWideEqualExpectedCount := 0;
        FNoneExpectedResult := E_Result.Passed;
        FNoneExpectedFinding := FALSE;
        FNoneExpectedCount := 0;
        FWideRangeExpectedResult := E_Result.Passed;
        FWideRangeExpectedFinding := FALSE;
        FWideRangeExpectedCount := 0;
    ScenarioFailedCount:
        FExpected := 3;
        FMinimum := 3;
        FMaximum := 3;
        FEqualExpectedResult := E_Result.Failed;
        FEqualExpectedFinding := TRUE;
        FEqualExpectedCount := 2;
        FWideEqualExpectedResult := E_Result.Failed;
        FWideEqualExpectedFinding := TRUE;
        FWideEqualExpectedCount := 2;
        FNoneExpectedResult := E_Result.Failed;
        FNoneExpectedFinding := TRUE;
        FNoneExpectedCount := 2;
        FWideRangeExpectedResult := E_Result.Failed;
        FWideRangeExpectedFinding := TRUE;
        FWideRangeExpectedCount := 2;
    ScenarioDisabledRetention:
        FContinueScenario := TRUE;
        FSubjectEnable := FALSE;
        FToken := 0;
        FWideToken := 0;
        FEqualExpectedResult := E_Result.Failed;
        FEqualExpectedFinding := FALSE;
        FEqualExpectedCount := 2;
        FWideEqualExpectedResult := E_Result.Failed;
        FWideEqualExpectedFinding := FALSE;
        FWideEqualExpectedCount := 2;
        FNoneExpectedResult := E_Result.Failed;
        FNoneExpectedFinding := FALSE;
        FNoneExpectedCount := 2;
        FWideRangeExpectedResult := E_Result.Failed;
        FWideRangeExpectedFinding := FALSE;
        FWideRangeExpectedCount := 2;
    ScenarioFailedRetention:
        FContinueScenario := TRUE;
        FToken := 0;
        FWideToken := 0;
        FEqualExpectedResult := E_Result.Failed;
        FEqualExpectedFinding := FALSE;
        FEqualExpectedCount := 2;
        FWideEqualExpectedResult := E_Result.Failed;
        FWideEqualExpectedFinding := FALSE;
        FWideEqualExpectedCount := 2;
        FNoneExpectedResult := E_Result.Failed;
        FNoneExpectedFinding := FALSE;
        FNoneExpectedCount := 2;
        FWideRangeExpectedResult := E_Result.Failed;
        FWideRangeExpectedFinding := FALSE;
        FWideRangeExpectedCount := 2;
    ScenarioErrorClearsCount:
        FContinueScenario := TRUE;
        FLength := 0;
        FEqualExpectedResult := E_Result.Error;
        FEqualExpectedFinding := TRUE;
        FEqualExpectedCount := 0;
        FWideEqualExpectedResult := E_Result.Error;
        FWideEqualExpectedFinding := TRUE;
        FWideEqualExpectedCount := 0;
        FNoneExpectedResult := E_Result.Error;
        FNoneExpectedFinding := TRUE;
        FNoneExpectedCount := 0;
        FWideRangeExpectedResult := E_Result.Error;
        FWideRangeExpectedFinding := TRUE;
        FWideRangeExpectedCount := 0;
    ScenarioResetAfterError:
        FEqualExpectedResult := E_Result.Passed;
        FEqualExpectedFinding := FALSE;
        FEqualExpectedCount := 2;
        FWideEqualExpectedResult := E_Result.Passed;
        FWideEqualExpectedFinding := FALSE;
        FWideEqualExpectedCount := 2;
        FNoneExpectedResult := E_Result.Failed;
        FNoneExpectedFinding := TRUE;
        FNoneExpectedCount := 2;
        FWideRangeExpectedResult := E_Result.Passed;
        FWideRangeExpectedFinding := FALSE;
        FWideRangeExpectedCount := 2;
    ScenarioBelowArray:
        FStartIndex := -3;
        FEqualExpectedResult := E_Result.Error;
        FEqualExpectedFinding := TRUE;
        FEqualExpectedCount := 0;
        FWideEqualExpectedResult := E_Result.Error;
        FWideEqualExpectedFinding := TRUE;
        FWideEqualExpectedCount := 0;
        FNoneExpectedResult := E_Result.Error;
        FNoneExpectedFinding := TRUE;
        FNoneExpectedCount := 0;
        FWideRangeExpectedResult := E_Result.Error;
        FWideRangeExpectedFinding := TRUE;
        FWideRangeExpectedCount := 0;
    ScenarioEndOutsideArray:
        FStartIndex := DINT#2147483647;
        FLength := 2;
        FEqualExpectedResult := E_Result.Error;
        FEqualExpectedFinding := TRUE;
        FEqualExpectedCount := 0;
        FWideEqualExpectedResult := E_Result.Error;
        FWideEqualExpectedFinding := TRUE;
        FWideEqualExpectedCount := 0;
        FNoneExpectedResult := E_Result.Error;
        FNoneExpectedFinding := TRUE;
        FNoneExpectedCount := 0;
        FWideRangeExpectedResult := E_Result.Error;
        FWideRangeExpectedFinding := TRUE;
        FWideRangeExpectedCount := 0;
    ScenarioReversedCountBounds:
        FMinimum := 3;
        FMaximum := 1;
        FEqualExpectedResult := E_Result.Passed;
        FEqualExpectedFinding := FALSE;
        FEqualExpectedCount := 2;
        FWideEqualExpectedResult := E_Result.Passed;
        FWideEqualExpectedFinding := FALSE;
        FWideEqualExpectedCount := 2;
        FNoneExpectedResult := E_Result.Failed;
        FNoneExpectedFinding := TRUE;
        FNoneExpectedCount := 2;
        FWideRangeExpectedResult := E_Result.Error;
        FWideRangeExpectedFinding := TRUE;
        FWideRangeExpectedCount := 0;
ELSE
    Error(Message := 'Unknown Assertion scenario.');
    RETURN;
END_CASE;
SelectScenario := TRUE;
END_METHOD

END_FUNCTION_BLOCK

// ---- SelfTests/TestCases/TestSuite_AssertionText/Test_AssertionArrayTokenCount.TcPOU
{region 'Documentation'}
(*!
<summary>Checks non-overlapping BYTE/WORD array token counts and independent array bounds.</summary>
<description>
Adjacent tokens count separately; overlapping candidates do not share elements.
Word patterns deliberately contain equal low bytes with different high bytes.
Oversized tokens and empty selected ranges are normal parameter errors, not
manufactured empty arrays or invalid references.
Independent scenarios occupy two calls: bound Reset, then evaluation.
ProcessAssertions checks each call before ProcessTests advances. Literal expected
results belong to SelectScenario, not to a copy of the production comparison.
The local capture is cleared before each call and checked in subject-call order.
FirstFailedScenario and FailedDuringEvaluation retain the first mismatch.
Continuation scenarios explicitly retain the prior subject state. The Test Case
owns all input storage; no invalid or dangling references are constructed.
</description>
*)
{endregion}
FUNCTION_BLOCK Test_AssertionArrayTokenCount EXTENDS TestCaseBase
VAR
    FEqual : AssertArrayTokenCntEqual_Byte;
    FEqualExpectedResult : E_Result;
    FWideEqual : AssertArrayTokenCntEqual_Word;
    FWideEqualExpectedResult : E_Result;
    FNone : AssertNoArrayToken_Byte;
    FNoneExpectedResult : E_Result;
    FWideRange : AssertArrayTokenCntInRange_Word;
    FWideRangeExpectedResult : E_Result;
    FData : ARRAY[-2..3] OF BYTE;
    FDataBefore : ARRAY[-2..3] OF BYTE;
    FWideData : ARRAY[-2..3] OF WORD;
    FWideDataBefore : ARRAY[-2..3] OF WORD;
    FToken : ARRAY[4..5] OF BYTE;
    FTokenBefore : ARRAY[4..5] OF BYTE;
    FWideToken : ARRAY[-5..-4] OF WORD;
    FWideTokenBefore : ARRAY[-5..-4] OF WORD;
    FStartIndex : DINT;
    FLength : USINT;
    FExpected : UINT;
    FMinimum : UINT;
    FMaximum : UINT;
    FSubjectEnable : BOOL;
    FContinueScenario : BOOL;
    FEqualExpectedFinding : BOOL;
    FEqualExpectedCount : UINT;
    FWideEqualExpectedFinding : BOOL;
    FWideEqualExpectedCount : UINT;
    FNoneExpectedFinding : BOOL;
    FNoneExpectedCount : UINT;
    FWideRangeExpectedFinding : BOOL;
    FWideRangeExpectedCount : UINT;
    FCapture : EventBuffer;
    FEvents : ARRAY[1..CaptureLength] OF ST_Event;
    FCaptureFifo : ST_FifoStatus;
    FCaptureStatus : ST_EventBufferStatus;
    FSetupValid : BOOL;
    FScenario : UINT;
    FChecked : BOOL;
    FEvaluateSubjects : BOOL;
    FObservationReady : BOOL;
    FFirstFailedScenario : UINT;
    FFailedDuringEvaluation : BOOL;
    FResultsMatch : BOOL;
    FResults : AssertTrue;
    FActivityMatch : BOOL;
    FActivity : AssertTrue;
    FInputsMatch : BOOL;
    FInputs : AssertTrue;
    FFindingsMatch : BOOL;
    FFindings : AssertTrue;
END_VAR
VAR CONSTANT
    CaptureLength : UINT := 8;
    ScenarioAdjacentTokens : UINT := 1;
    ScenarioNonOverlapping : UINT := 2;
    ScenarioTrailingPartial : UINT := 3;
    ScenarioLastCandidate : UINT := 4;
    ScenarioAbsent : UINT := 5;
    ScenarioCountMismatch : UINT := 6;
    ScenarioTokenTooLong : UINT := 7;
    ScenarioEmptyRange : UINT := 8;
    ScenarioRangePastEnd : UINT := 9;
    LastScenario : UINT := ScenarioRangePastEnd;
END_VAR

SUPER^();

{region 'Documentation'}
(*!
<summary>Aggregates only outer checks, not intentionally failing subjects.</summary>
*)
{endregion}
METHOD PROTECTED AggregateResults
VAR_INPUT
    Aggregator : I_ResultAggregator; //! Borrowed result sink owned by the outer Test Case; add this test's checking Assertions without resetting or retaining the sink.
END_VAR
Aggregator.AddProvider(Provider := FResults);
Aggregator.AddProvider(Provider := FActivity);
Aggregator.AddProvider(Provider := FInputs);
Aggregator.AddProvider(Provider := FFindings);
END_METHOD

{region 'Documentation'}
(*!
<summary>Calls each inherited production subject once with caller-owned input storage.</summary>
*)
{endregion}
METHOD PRIVATE CallSubjects
FEqual(Enable := FSubjectEnable,
    State := E_State.Running,
    StartIndex := FStartIndex,
    Length := FLength,
    Expected := FExpected,
    IN := FData,
    Token := FToken);
FWideEqual(Enable := FSubjectEnable,
    State := E_State.Running,
    StartIndex := FStartIndex,
    Length := FLength,
    Expected := FExpected,
    IN := FWideData,
    Token := FWideToken);
FNone(Enable := FSubjectEnable,
    State := E_State.Running,
    StartIndex := FStartIndex,
    Length := FLength,
    IN := FData,
    Token := FToken);
FWideRange(Enable := FSubjectEnable,
    State := E_State.Running,
    StartIndex := FStartIndex,
    Length := FLength,
    Minimum := FMinimum,
    Maximum := FMaximum,
    IN := FWideData,
    Token := FWideToken);
END_METHOD

{region 'Documentation'}
(*!
<summary>Checks one subject finding in call order; expected outcomes come from the scenario.</summary>
*)
{endregion}
METHOD PRIVATE CheckFinding : BOOL //! TRUE when the required finding checks pass; calls requiring no finding also succeed.
VAR_INPUT
    Subject : I_Assertion; //! Assertion interface supplying the expected finding identity.
    ExpectedResult : E_Result; //! Independently authored result expected in the captured finding.
    ExpectedFinding : BOOL; //! TRUE when this scenario requires a finding during active evaluation.
END_VAR
VAR_IN_OUT
    Index : UINT; //! One-based next finding index; advanced when this call checks a required finding.
END_VAR
CheckFinding := TRUE;
IF FEvaluateSubjects AND ExpectedFinding THEN
    CheckFinding := (FEvents[Index].SequenceId = UINT_TO_UDINT(Index))
        AND (FEvents[Index].Name = Subject.Name)
        AND (FEvents[Index].OwnerScope = E_OwnerScope.Assertion)
        AND (FEvents[Index].EventType = E_EventType.Result)
        AND (FEvents[Index].State = E_State.Running)
        AND (FEvents[Index].Result = ExpectedResult)
        AND (FEvents[Index].Message <> '');
    Index := Index + 1;
END_IF;
END_METHOD

{region 'Documentation'}
(*!
<summary>Checks exact finding count and identities; at most one finding per subject.</summary>
*)
{endregion}
METHOD PRIVATE CheckFindings
VAR
    Index : UINT;
    Matches : BOOL;
END_VAR
Index := 1;
FFindingsMatch := TRUE;
Matches := CheckFinding(Subject := FEqual,
    ExpectedResult := FEqualExpectedResult,
    ExpectedFinding := FEqualExpectedFinding,
    Index := Index);
FFindingsMatch := FFindingsMatch AND Matches;
Matches := CheckFinding(Subject := FWideEqual,
    ExpectedResult := FWideEqualExpectedResult,
    ExpectedFinding := FWideEqualExpectedFinding,
    Index := Index);
FFindingsMatch := FFindingsMatch AND Matches;
Matches := CheckFinding(Subject := FNone,
    ExpectedResult := FNoneExpectedResult,
    ExpectedFinding := FNoneExpectedFinding,
    Index := Index);
FFindingsMatch := FFindingsMatch AND Matches;
Matches := CheckFinding(Subject := FWideRange,
    ExpectedResult := FWideRangeExpectedResult,
    ExpectedFinding := FWideRangeExpectedFinding,
    Index := Index);
FFindingsMatch := FFindingsMatch AND Matches;
FFindingsMatch := FFindingsMatch
    AND (FCaptureStatus.SequenceId = UINT_TO_UDINT(Index - 1))
    AND (FCaptureStatus.LostEventCount = 0);
IF FEvaluateSubjects AND (FScenario = ScenarioCountMismatch) THEN
    // SA0175: Fixed byte-substring checks of bounded diagnostic messages; no character offsets.
    {analysis -175}
    FFindingsMatch := FFindingsMatch
        AND (FIND(FEvents[1].Message, 'Actual = 2') > 0)
        AND (FIND(FEvents[4].Message, 'Actual = 2') > 0);
    {analysis +175}
END_IF;
END_METHOD

{region 'Documentation'}
(*!
<summary>Rejects incomplete subject, capture or outer Assertion setup.</summary>
*)
{endregion}
METHOD PROTECTED CheckInitialization : BOOL //! TRUE when the inherited initialization check and this concrete fixture check both accept the setup.
CheckInitialization := SUPER^.CheckInitialization();
IF NOT CheckInitialization THEN
    RETURN;
END_IF;

CheckInitialization := FSetupValid
    AND FResults.IsInitialized
    AND FActivity.IsInitialized
    AND FInputs.IsInitialized
    AND FFindings.IsInitialized;
IF NOT CheckInitialization THEN
    EventPublisher.PublishEvent(Event := CreateFrameworkEvent(Name := Name,
        ResourceName := '',
        State := State,
        Severity := E_EventSeverity.Error,
        Message := 'Text selftest setup failed.'));
END_IF;
END_METHOD

{region 'Documentation'}
(*!
<summary>Checks literal evaluation results, or NotEvaluated on the reset call.</summary>
*)
{endregion}
METHOD PRIVATE CheckResults
IF FEvaluateSubjects THEN
    FResultsMatch := (FEqual.Result = FEqualExpectedResult)
        AND (FWideEqual.Result = FWideEqualExpectedResult)
        AND (FNone.Result = FNoneExpectedResult)
        AND (FWideRange.Result = FWideRangeExpectedResult);
ELSE
    FResultsMatch := (FEqual.Result = E_Result.NotEvaluated)
        AND (FWideEqual.Result = E_Result.NotEvaluated)
        AND (FNone.Result = E_Result.NotEvaluated)
        AND (FWideRange.Result = E_Result.NotEvaluated);
END_IF;
FActivityMatch := (FEqual.Enabled = FSubjectEnable)
    AND (FEqual.ObservationActive = (FEvaluateSubjects AND FSubjectEnable))
    AND (FEqual.EvaluationActive = (FEvaluateSubjects AND FSubjectEnable))
    AND (FWideEqual.Enabled = FSubjectEnable)
    AND (FWideEqual.ObservationActive = (FEvaluateSubjects AND FSubjectEnable))
    AND (FWideEqual.EvaluationActive = (FEvaluateSubjects AND FSubjectEnable))
    AND (FNone.Enabled = FSubjectEnable)
    AND (FNone.ObservationActive = (FEvaluateSubjects AND FSubjectEnable))
    AND (FNone.EvaluationActive = (FEvaluateSubjects AND FSubjectEnable))
    AND (FWideRange.Enabled = FSubjectEnable)
    AND (FWideRange.ObservationActive = (FEvaluateSubjects AND FSubjectEnable))
    AND (FWideRange.EvaluationActive = (FEvaluateSubjects AND FSubjectEnable));
IF FEvaluateSubjects THEN
    FResultsMatch := FResultsMatch
        AND (FEqual.TokenCount = FEqualExpectedCount)
        AND (FWideEqual.TokenCount = FWideEqualExpectedCount)
        AND (FNone.TokenCount = FNoneExpectedCount)
        AND (FWideRange.TokenCount = FWideRangeExpectedCount);
ELSE
    FResultsMatch := FResultsMatch
        AND (FEqual.TokenCount = 0)
        AND (FWideEqual.TokenCount = 0)
        AND (FNone.TokenCount = 0)
        AND (FWideRange.TokenCount = 0);
END_IF;
END_METHOD

{region 'Documentation'}
(*!
<summary>Initializes outer checks and isolates intentional subject findings.</summary>
*)
{endregion}
METHOD PROTECTED Configure
VAR
    Initialized : BOOL;
END_VAR
FPreparationStateCount := 0;
FTestStateCount := 1;
FResults.Initialize(Parent := THIS^,
    AssertionName := 'Results');
FActivity.Initialize(Parent := THIS^,
    AssertionName := 'Activity');
FInputs.Initialize(Parent := THIS^,
    AssertionName := 'Inputs');
FFindings.Initialize(Parent := THIS^,
    AssertionName := 'Findings');
FSetupValid := FCapture.Initialize(Buffer := FEvents,
    FifoControl := FCaptureFifo,
    Status := FCaptureStatus);
FEqual.BindPublisher(Publisher := FCapture);
Initialized := FEqual.Initialize(Parent := THIS^,
    AssertionName := 'Equal');
FSetupValid := FSetupValid AND Initialized;
FWideEqual.BindPublisher(Publisher := FCapture);
Initialized := FWideEqual.Initialize(Parent := THIS^,
    AssertionName := 'WideEqual');
FSetupValid := FSetupValid AND Initialized;
FNone.BindPublisher(Publisher := FCapture);
Initialized := FNone.Initialize(Parent := THIS^,
    AssertionName := 'None');
FSetupValid := FSetupValid AND Initialized;
FWideRange.BindPublisher(Publisher := FCapture);
Initialized := FWideRange.Initialize(Parent := THIS^,
    AssertionName := 'WideRange');
FSetupValid := FSetupValid AND Initialized;
END_METHOD

{region 'Documentation'}
(*!
<summary>Completes abort; no asynchronous resource is owned.</summary>
*)
{endregion}
METHOD PROTECTED ProcessAbort
VAR_INPUT
    Enable : BOOL; //! Phase permission supplied by the owning Test Case; FALSE does not authorize progression, while observation may continue.
END_VAR
IF Enable THEN
    CompleteAbort();
END_IF;
END_METHOD

{region 'Documentation'}
(*!
<summary>Latches this call's checks before progression is permitted.</summary>
*)
{endregion}
METHOD PROTECTED ProcessAssertions
VAR_INPUT
    Enable : BOOL; //! Phase permission supplied by the owning Test Case; FALSE does not authorize progression, while observation may continue.
END_VAR
VAR
    Check : BOOL;
END_VAR
Check := Enable AND FObservationReady;
FResults(Enable := Check,
    State := State,
    IN := FResultsMatch);
FActivity(Enable := Check,
    State := State,
    IN := FActivityMatch);
FInputs(Enable := Check,
    State := State,
    IN := FInputsMatch);
FFindings(Enable := Check,
    State := State,
    IN := FFindingsMatch);
IF Check THEN
    FChecked := TRUE;
END_IF;
END_METHOD

{region 'Documentation'}
(*!
<summary>No Preparation phase is needed.</summary>
*)
{endregion}
METHOD PROTECTED ProcessPreparations
VAR_INPUT
    // SA0033: Required hook; this test has no Preparation phase.
    {attribute 'analysis' := '-33'}
    Enable : BOOL; //! Phase permission supplied by the owning Test Case; FALSE does not authorize progression, while observation may continue.
END_VAR
END_METHOD

{region 'Documentation'}
(*!
<summary>Restarts the scenario sequence and outer checks.</summary>
*)
{endregion}
METHOD PROTECTED ProcessReset
FScenario := ScenarioAdjacentTokens;
FChecked := FALSE;
FSubjectEnable := FALSE;
FContinueScenario := FALSE;
FEvaluateSubjects := FALSE;
FObservationReady := FALSE;
FFirstFailedScenario := 0;
FFailedDuringEvaluation := FALSE;
FCapture.Reset();
ResetSubjects();
FResults.Reset();
FActivity.Reset();
FInputs.Reset();
FFindings.Reset();
CompleteReset();
END_METHOD

{region 'Documentation'}
(*!
<summary>Consumes reset before each independent scenario; continuation retains subject state.</summary>
*)
{endregion}
METHOD PROTECTED ProcessTests
VAR_INPUT
    Enable : BOOL; //! Phase permission supplied by the owning Test Case; FALSE does not authorize progression, while observation may continue.
END_VAR
IF NOT Enable THEN
    RETURN;
END_IF;

IF FChecked THEN
    FChecked := FALSE;
    FObservationReady := FALSE;
    IF FEvaluateSubjects THEN
        IF FScenario = LastScenario THEN
            CompleteTests();
            RETURN;
        END_IF;
        FScenario := FScenario + 1;
    END_IF;
    FEvaluateSubjects := NOT FEvaluateSubjects;
END_IF;

IF NOT SelectScenario() THEN
    RETURN;
END_IF;
IF FContinueScenario THEN
    FEvaluateSubjects := TRUE;
END_IF;
FCapture.Reset();
IF NOT FEvaluateSubjects THEN
    ResetSubjects();
END_IF;
FDataBefore := FData;
FWideDataBefore := FWideData;
FTokenBefore := FToken;
FWideTokenBefore := FWideToken;
CallSubjects();
CheckResults();
FInputsMatch := (FData[-2] = FDataBefore[-2])
    AND (FData[-1] = FDataBefore[-1])
    AND (FData[0] = FDataBefore[0])
    AND (FData[1] = FDataBefore[1])
    AND (FData[2] = FDataBefore[2])
    AND (FData[3] = FDataBefore[3])
    AND (FWideData[-2] = FWideDataBefore[-2])
    AND (FWideData[-1] = FWideDataBefore[-1])
    AND (FWideData[0] = FWideDataBefore[0])
    AND (FWideData[1] = FWideDataBefore[1])
    AND (FWideData[2] = FWideDataBefore[2])
    AND (FWideData[3] = FWideDataBefore[3])
    AND (FToken[4] = FTokenBefore[4])
    AND (FToken[5] = FTokenBefore[5])
    AND (FWideToken[-5] = FWideTokenBefore[-5])
    AND (FWideToken[-4] = FWideTokenBefore[-4]);
CheckFindings();
IF (FFirstFailedScenario = 0)
    AND NOT (FResultsMatch AND FActivityMatch AND FInputsMatch AND FFindingsMatch) THEN
    FFirstFailedScenario := FScenario;
    FFailedDuringEvaluation := FEvaluateSubjects;
END_IF;
FObservationReady := TRUE;
END_METHOD

{region 'Documentation'}
(*!
<summary>Queues reset; the next bound FB call consumes it without evaluating.</summary>
*)
{endregion}
METHOD PRIVATE ResetSubjects
FEqual.Reset();
FWideEqual.Reset();
FNone.Reset();
FWideRange.Reset();
END_METHOD

{region 'Documentation'}
(*!
<summary>Selects explicit stimuli and expected results for one scenario.</summary>
*)
{endregion}
METHOD PRIVATE SelectScenario : BOOL //! TRUE after selecting a supported scenario and its literal expectations; FALSE reports an unknown scenario.
SelectScenario := FALSE;
FSubjectEnable := TRUE;
FContinueScenario := FALSE;
FData[-2] := 1;
FData[-1] := 2;
FData[0] := 1;
FData[1] := 2;
FData[2] := 9;
FData[3] := 9;
FWideData[-2] := WORD#16#0101;
FWideData[-1] := WORD#16#0202;
FWideData[0] := WORD#16#0101;
FWideData[1] := WORD#16#0202;
FWideData[2] := 1;
FWideData[3] := 2;
FToken[4] := 1;
FToken[5] := 2;
FWideToken[-5] := WORD#16#0101;
FWideToken[-4] := WORD#16#0202;
FStartIndex := -2;
FLength := 6;
FExpected := 2;
FMinimum := 2;
FMaximum := 2;
CASE FScenario OF
    ScenarioAdjacentTokens:
        FEqualExpectedResult := E_Result.Passed;
        FEqualExpectedFinding := FALSE;
        FEqualExpectedCount := 2;
        FWideEqualExpectedResult := E_Result.Passed;
        FWideEqualExpectedFinding := FALSE;
        FWideEqualExpectedCount := 2;
        FNoneExpectedResult := E_Result.Failed;
        FNoneExpectedFinding := TRUE;
        FNoneExpectedCount := 2;
        FWideRangeExpectedResult := E_Result.Passed;
        FWideRangeExpectedFinding := FALSE;
        FWideRangeExpectedCount := 2;
    ScenarioNonOverlapping:
        FLength := 3;
        FData[-1] := 1;
        FToken[5] := 1;
        FWideData[-1] := WORD#16#0101;
        FWideToken[-4] := WORD#16#0101;
        FExpected := 1;
        FMinimum := 1;
        FMaximum := 1;
        FEqualExpectedResult := E_Result.Passed;
        FEqualExpectedFinding := FALSE;
        FEqualExpectedCount := 1;
        FWideEqualExpectedResult := E_Result.Passed;
        FWideEqualExpectedFinding := FALSE;
        FWideEqualExpectedCount := 1;
        FNoneExpectedResult := E_Result.Failed;
        FNoneExpectedFinding := TRUE;
        FNoneExpectedCount := 1;
        FWideRangeExpectedResult := E_Result.Passed;
        FWideRangeExpectedFinding := FALSE;
        FWideRangeExpectedCount := 1;
    ScenarioTrailingPartial:
        FLength := 3;
        FExpected := 1;
        FMinimum := 1;
        FMaximum := 1;
        FEqualExpectedResult := E_Result.Passed;
        FEqualExpectedFinding := FALSE;
        FEqualExpectedCount := 1;
        FWideEqualExpectedResult := E_Result.Passed;
        FWideEqualExpectedFinding := FALSE;
        FWideEqualExpectedCount := 1;
        FNoneExpectedResult := E_Result.Failed;
        FNoneExpectedFinding := TRUE;
        FNoneExpectedCount := 1;
        FWideRangeExpectedResult := E_Result.Passed;
        FWideRangeExpectedFinding := FALSE;
        FWideRangeExpectedCount := 1;
    ScenarioLastCandidate:
        FStartIndex := -1;
        FLength := 3;
        FExpected := 1;
        FMinimum := 1;
        FMaximum := 1;
        FEqualExpectedResult := E_Result.Passed;
        FEqualExpectedFinding := FALSE;
        FEqualExpectedCount := 1;
        FWideEqualExpectedResult := E_Result.Passed;
        FWideEqualExpectedFinding := FALSE;
        FWideEqualExpectedCount := 1;
        FNoneExpectedResult := E_Result.Failed;
        FNoneExpectedFinding := TRUE;
        FNoneExpectedCount := 1;
        FWideRangeExpectedResult := E_Result.Passed;
        FWideRangeExpectedFinding := FALSE;
        FWideRangeExpectedCount := 1;
    ScenarioAbsent:
        FToken[4] := 7;
        FWideToken[-5] := 7;
        FExpected := 0;
        FMinimum := 0;
        FMaximum := 0;
        FEqualExpectedResult := E_Result.Passed;
        FEqualExpectedFinding := FALSE;
        FEqualExpectedCount := 0;
        FWideEqualExpectedResult := E_Result.Passed;
        FWideEqualExpectedFinding := FALSE;
        FWideEqualExpectedCount := 0;
        FNoneExpectedResult := E_Result.Passed;
        FNoneExpectedFinding := FALSE;
        FNoneExpectedCount := 0;
        FWideRangeExpectedResult := E_Result.Passed;
        FWideRangeExpectedFinding := FALSE;
        FWideRangeExpectedCount := 0;
    ScenarioCountMismatch:
        FExpected := 1;
        FMinimum := 3;
        FMaximum := 4;
        FEqualExpectedResult := E_Result.Failed;
        FEqualExpectedFinding := TRUE;
        FEqualExpectedCount := 2;
        FWideEqualExpectedResult := E_Result.Failed;
        FWideEqualExpectedFinding := TRUE;
        FWideEqualExpectedCount := 2;
        FNoneExpectedResult := E_Result.Failed;
        FNoneExpectedFinding := TRUE;
        FNoneExpectedCount := 2;
        FWideRangeExpectedResult := E_Result.Failed;
        FWideRangeExpectedFinding := TRUE;
        FWideRangeExpectedCount := 2;
    ScenarioTokenTooLong:
        FLength := 1;
        FEqualExpectedResult := E_Result.Error;
        FEqualExpectedFinding := TRUE;
        FEqualExpectedCount := 0;
        FWideEqualExpectedResult := E_Result.Error;
        FWideEqualExpectedFinding := TRUE;
        FWideEqualExpectedCount := 0;
        FNoneExpectedResult := E_Result.Error;
        FNoneExpectedFinding := TRUE;
        FNoneExpectedCount := 0;
        FWideRangeExpectedResult := E_Result.Error;
        FWideRangeExpectedFinding := TRUE;
        FWideRangeExpectedCount := 0;
    ScenarioEmptyRange:
        FLength := 0;
        FEqualExpectedResult := E_Result.Error;
        FEqualExpectedFinding := TRUE;
        FEqualExpectedCount := 0;
        FWideEqualExpectedResult := E_Result.Error;
        FWideEqualExpectedFinding := TRUE;
        FWideEqualExpectedCount := 0;
        FNoneExpectedResult := E_Result.Error;
        FNoneExpectedFinding := TRUE;
        FNoneExpectedCount := 0;
        FWideRangeExpectedResult := E_Result.Error;
        FWideRangeExpectedFinding := TRUE;
        FWideRangeExpectedCount := 0;
    ScenarioRangePastEnd:
        FStartIndex := 3;
        FLength := 2;
        FEqualExpectedResult := E_Result.Error;
        FEqualExpectedFinding := TRUE;
        FEqualExpectedCount := 0;
        FWideEqualExpectedResult := E_Result.Error;
        FWideEqualExpectedFinding := TRUE;
        FWideEqualExpectedCount := 0;
        FNoneExpectedResult := E_Result.Error;
        FNoneExpectedFinding := TRUE;
        FNoneExpectedCount := 0;
        FWideRangeExpectedResult := E_Result.Error;
        FWideRangeExpectedFinding := TRUE;
        FWideRangeExpectedCount := 0;
ELSE
    Error(Message := 'Unknown Assertion scenario.');
    RETURN;
END_CASE;
SelectScenario := TRUE;
END_METHOD

END_FUNCTION_BLOCK

// ---- SelfTests/TestCases/TestSuite_AssertionText/Test_AssertionLengthUntil.TcPOU
{region 'Documentation'}
(*!
<summary>Checks first-token distance in elements for BYTE/WORD value and array tokens.</summary>
<description>
The first matching index is measured relative to StartIndex, excluding the token.
No match is Failed even for NotEqual. Array bounds are independent of the token
bounds; Word data makes element distance distinguishable from byte distance.
Independent scenarios occupy two calls: bound Reset, then evaluation.
ProcessAssertions checks each call before ProcessTests advances. Literal expected
results belong to SelectScenario, not to a copy of the production comparison.
The local capture is cleared before each call and checked in subject-call order.
FirstFailedScenario and FailedDuringEvaluation retain the first mismatch.
Continuation scenarios explicitly retain the prior subject state. The Test Case
owns all input storage; no invalid or dangling references are constructed.
</description>
*)
{endregion}
FUNCTION_BLOCK Test_AssertionLengthUntil EXTENDS TestCaseBase
VAR
    FValue : AssertLengthUntilValueEqual_Byte;
    FValueExpectedResult : E_Result;
    FWideValue : AssertLengthUntilValueNotEqual_Word;
    FWideValueExpectedResult : E_Result;
    FArray : AssertLengthUntilArrayNotEqual_Byte;
    FArrayExpectedResult : E_Result;
    FWideArray : AssertLengthUntilArrayEqual_Word;
    FWideArrayExpectedResult : E_Result;
    FData : ARRAY[-2..3] OF BYTE;
    FDataBefore : ARRAY[-2..3] OF BYTE;
    FWideData : ARRAY[-2..3] OF WORD;
    FWideDataBefore : ARRAY[-2..3] OF WORD;
    FToken : ARRAY[4..5] OF BYTE;
    FTokenBefore : ARRAY[4..5] OF BYTE;
    FWideToken : ARRAY[-5..-4] OF WORD;
    FWideTokenBefore : ARRAY[-5..-4] OF WORD;
    FStartIndex : DINT;
    FLength : USINT;
    FExpected : USINT;
    FValueToken : BYTE;
    FWideValueToken : WORD;
    FMask : BYTE;
    FWideMask : WORD;
    FSubjectEnable : BOOL;
    FContinueScenario : BOOL;
    FValueExpectedFinding : BOOL;
    FWideValueExpectedFinding : BOOL;
    FArrayExpectedFinding : BOOL;
    FWideArrayExpectedFinding : BOOL;
    FCapture : EventBuffer;
    FEvents : ARRAY[1..CaptureLength] OF ST_Event;
    FCaptureFifo : ST_FifoStatus;
    FCaptureStatus : ST_EventBufferStatus;
    FSetupValid : BOOL;
    FScenario : UINT;
    FChecked : BOOL;
    FEvaluateSubjects : BOOL;
    FObservationReady : BOOL;
    FFirstFailedScenario : UINT;
    FFailedDuringEvaluation : BOOL;
    FResultsMatch : BOOL;
    FResults : AssertTrue;
    FActivityMatch : BOOL;
    FActivity : AssertTrue;
    FInputsMatch : BOOL;
    FInputs : AssertTrue;
    FFindingsMatch : BOOL;
    FFindings : AssertTrue;
END_VAR
VAR CONSTANT
    CaptureLength : UINT := 8;
    ScenarioFirstOfMultiple : UINT := 1;
    ScenarioAtStart : UINT := 2;
    ScenarioLastCandidate : UINT := 3;
    ScenarioDistanceMismatch : UINT := 4;
    ScenarioElementDistance : UINT := 5;
    ScenarioMaskedValue : UINT := 6;
    ScenarioLastValue : UINT := 7;
    ScenarioAbsent : UINT := 8;
    ScenarioTokenTooLong : UINT := 9;
    ScenarioEmptyRange : UINT := 10;
    ScenarioRangePastEnd : UINT := 11;
    LastScenario : UINT := ScenarioRangePastEnd;
END_VAR

SUPER^();

{region 'Documentation'}
(*!
<summary>Aggregates only outer checks, not intentionally failing subjects.</summary>
*)
{endregion}
METHOD PROTECTED AggregateResults
VAR_INPUT
    Aggregator : I_ResultAggregator; //! Borrowed result sink owned by the outer Test Case; add this test's checking Assertions without resetting or retaining the sink.
END_VAR
Aggregator.AddProvider(Provider := FResults);
Aggregator.AddProvider(Provider := FActivity);
Aggregator.AddProvider(Provider := FInputs);
Aggregator.AddProvider(Provider := FFindings);
END_METHOD

{region 'Documentation'}
(*!
<summary>Calls each inherited production subject once with caller-owned input storage.</summary>
*)
{endregion}
METHOD PRIVATE CallSubjects
FValue(Enable := FSubjectEnable,
    State := E_State.Running,
    StartIndex := FStartIndex,
    Length := FLength,
    Expected := FExpected,
    Token := FValueToken,
    Mask := FMask,
    IN := FData);
FWideValue(Enable := FSubjectEnable,
    State := E_State.Running,
    StartIndex := FStartIndex,
    Length := FLength,
    Expected := FExpected,
    Token := FWideValueToken,
    Mask := FWideMask,
    IN := FWideData);
FArray(Enable := FSubjectEnable,
    State := E_State.Running,
    StartIndex := FStartIndex,
    Length := FLength,
    Expected := FExpected,
    Token := FToken,
    IN := FData);
FWideArray(Enable := FSubjectEnable,
    State := E_State.Running,
    StartIndex := FStartIndex,
    Length := FLength,
    Expected := FExpected,
    Token := FWideToken,
    IN := FWideData);
END_METHOD

{region 'Documentation'}
(*!
<summary>Checks one subject finding in call order; expected outcomes come from the scenario.</summary>
*)
{endregion}
METHOD PRIVATE CheckFinding : BOOL //! TRUE when the required finding checks pass; calls requiring no finding also succeed.
VAR_INPUT
    Subject : I_Assertion; //! Assertion interface supplying the expected finding identity.
    ExpectedResult : E_Result; //! Independently authored result expected in the captured finding.
    ExpectedFinding : BOOL; //! TRUE when this scenario requires a finding during active evaluation.
END_VAR
VAR_IN_OUT
    Index : UINT; //! One-based next finding index; advanced when this call checks a required finding.
END_VAR
CheckFinding := TRUE;
IF FEvaluateSubjects AND ExpectedFinding THEN
    CheckFinding := (FEvents[Index].SequenceId = UINT_TO_UDINT(Index))
        AND (FEvents[Index].Name = Subject.Name)
        AND (FEvents[Index].OwnerScope = E_OwnerScope.Assertion)
        AND (FEvents[Index].EventType = E_EventType.Result)
        AND (FEvents[Index].State = E_State.Running)
        AND (FEvents[Index].Result = ExpectedResult)
        AND (FEvents[Index].Message <> '');
    Index := Index + 1;
END_IF;
END_METHOD

{region 'Documentation'}
(*!
<summary>Checks exact finding count and identities; at most one finding per subject.</summary>
*)
{endregion}
METHOD PRIVATE CheckFindings
VAR
    Index : UINT;
    Matches : BOOL;
END_VAR
Index := 1;
FFindingsMatch := TRUE;
Matches := CheckFinding(Subject := FValue,
    ExpectedResult := FValueExpectedResult,
    ExpectedFinding := FValueExpectedFinding,
    Index := Index);
FFindingsMatch := FFindingsMatch AND Matches;
Matches := CheckFinding(Subject := FWideValue,
    ExpectedResult := FWideValueExpectedResult,
    ExpectedFinding := FWideValueExpectedFinding,
    Index := Index);
FFindingsMatch := FFindingsMatch AND Matches;
Matches := CheckFinding(Subject := FArray,
    ExpectedResult := FArrayExpectedResult,
    ExpectedFinding := FArrayExpectedFinding,
    Index := Index);
FFindingsMatch := FFindingsMatch AND Matches;
Matches := CheckFinding(Subject := FWideArray,
    ExpectedResult := FWideArrayExpectedResult,
    ExpectedFinding := FWideArrayExpectedFinding,
    Index := Index);
FFindingsMatch := FFindingsMatch AND Matches;
FFindingsMatch := FFindingsMatch
    AND (FCaptureStatus.SequenceId = UINT_TO_UDINT(Index - 1))
    AND (FCaptureStatus.LostEventCount = 0);
IF FEvaluateSubjects AND (FScenario = ScenarioAbsent) THEN
    FFindingsMatch := FFindingsMatch
        AND (FEvents[1].Message = 'Assertion failed: token not found. StartIndex = -2, Length = 6')
        AND (FEvents[2].Message = FEvents[1].Message)
        AND (FEvents[3].Message = FEvents[1].Message)
        AND (FEvents[4].Message = FEvents[1].Message);
END_IF;
IF FEvaluateSubjects AND (FScenario = ScenarioDistanceMismatch) THEN
    // SA0175: Fixed byte-substring checks of bounded diagnostic messages; no character offsets.
    {analysis -175}
    FFindingsMatch := FFindingsMatch
        AND (FIND(FEvents[1].Message, 'Expected = 2, Actual = 1') > 0)
        AND (FIND(FEvents[2].Message, 'Expected = 2, Actual = 1') > 0);
    {analysis +175}
END_IF;
END_METHOD

{region 'Documentation'}
(*!
<summary>Rejects incomplete subject, capture or outer Assertion setup.</summary>
*)
{endregion}
METHOD PROTECTED CheckInitialization : BOOL //! TRUE when the inherited initialization check and this concrete fixture check both accept the setup.
CheckInitialization := SUPER^.CheckInitialization();
IF NOT CheckInitialization THEN
    RETURN;
END_IF;

CheckInitialization := FSetupValid
    AND FResults.IsInitialized
    AND FActivity.IsInitialized
    AND FInputs.IsInitialized
    AND FFindings.IsInitialized;
IF NOT CheckInitialization THEN
    EventPublisher.PublishEvent(Event := CreateFrameworkEvent(Name := Name,
        ResourceName := '',
        State := State,
        Severity := E_EventSeverity.Error,
        Message := 'Text selftest setup failed.'));
END_IF;
END_METHOD

{region 'Documentation'}
(*!
<summary>Checks literal evaluation results, or NotEvaluated on the reset call.</summary>
*)
{endregion}
METHOD PRIVATE CheckResults
IF FEvaluateSubjects THEN
    FResultsMatch := (FValue.Result = FValueExpectedResult)
        AND (FWideValue.Result = FWideValueExpectedResult)
        AND (FArray.Result = FArrayExpectedResult)
        AND (FWideArray.Result = FWideArrayExpectedResult);
ELSE
    FResultsMatch := (FValue.Result = E_Result.NotEvaluated)
        AND (FWideValue.Result = E_Result.NotEvaluated)
        AND (FArray.Result = E_Result.NotEvaluated)
        AND (FWideArray.Result = E_Result.NotEvaluated);
END_IF;
FActivityMatch := (FValue.Enabled = FSubjectEnable)
    AND (FValue.ObservationActive = (FEvaluateSubjects AND FSubjectEnable))
    AND (FValue.EvaluationActive = (FEvaluateSubjects AND FSubjectEnable))
    AND (FWideValue.Enabled = FSubjectEnable)
    AND (FWideValue.ObservationActive = (FEvaluateSubjects AND FSubjectEnable))
    AND (FWideValue.EvaluationActive = (FEvaluateSubjects AND FSubjectEnable))
    AND (FArray.Enabled = FSubjectEnable)
    AND (FArray.ObservationActive = (FEvaluateSubjects AND FSubjectEnable))
    AND (FArray.EvaluationActive = (FEvaluateSubjects AND FSubjectEnable))
    AND (FWideArray.Enabled = FSubjectEnable)
    AND (FWideArray.ObservationActive = (FEvaluateSubjects AND FSubjectEnable))
    AND (FWideArray.EvaluationActive = (FEvaluateSubjects AND FSubjectEnable));
END_METHOD

{region 'Documentation'}
(*!
<summary>Initializes outer checks and isolates intentional subject findings.</summary>
*)
{endregion}
METHOD PROTECTED Configure
VAR
    Initialized : BOOL;
END_VAR
FPreparationStateCount := 0;
FTestStateCount := 1;
FResults.Initialize(Parent := THIS^,
    AssertionName := 'Results');
FActivity.Initialize(Parent := THIS^,
    AssertionName := 'Activity');
FInputs.Initialize(Parent := THIS^,
    AssertionName := 'Inputs');
FFindings.Initialize(Parent := THIS^,
    AssertionName := 'Findings');
FSetupValid := FCapture.Initialize(Buffer := FEvents,
    FifoControl := FCaptureFifo,
    Status := FCaptureStatus);
FValue.BindPublisher(Publisher := FCapture);
Initialized := FValue.Initialize(Parent := THIS^,
    AssertionName := 'Value');
FSetupValid := FSetupValid AND Initialized;
FWideValue.BindPublisher(Publisher := FCapture);
Initialized := FWideValue.Initialize(Parent := THIS^,
    AssertionName := 'WideValue');
FSetupValid := FSetupValid AND Initialized;
FArray.BindPublisher(Publisher := FCapture);
Initialized := FArray.Initialize(Parent := THIS^,
    AssertionName := 'Array');
FSetupValid := FSetupValid AND Initialized;
FWideArray.BindPublisher(Publisher := FCapture);
Initialized := FWideArray.Initialize(Parent := THIS^,
    AssertionName := 'WideArray');
FSetupValid := FSetupValid AND Initialized;
END_METHOD

{region 'Documentation'}
(*!
<summary>Completes abort; no asynchronous resource is owned.</summary>
*)
{endregion}
METHOD PROTECTED ProcessAbort
VAR_INPUT
    Enable : BOOL; //! Phase permission supplied by the owning Test Case; FALSE does not authorize progression, while observation may continue.
END_VAR
IF Enable THEN
    CompleteAbort();
END_IF;
END_METHOD

{region 'Documentation'}
(*!
<summary>Latches this call's checks before progression is permitted.</summary>
*)
{endregion}
METHOD PROTECTED ProcessAssertions
VAR_INPUT
    Enable : BOOL; //! Phase permission supplied by the owning Test Case; FALSE does not authorize progression, while observation may continue.
END_VAR
VAR
    Check : BOOL;
END_VAR
Check := Enable AND FObservationReady;
FResults(Enable := Check,
    State := State,
    IN := FResultsMatch);
FActivity(Enable := Check,
    State := State,
    IN := FActivityMatch);
FInputs(Enable := Check,
    State := State,
    IN := FInputsMatch);
FFindings(Enable := Check,
    State := State,
    IN := FFindingsMatch);
IF Check THEN
    FChecked := TRUE;
END_IF;
END_METHOD

{region 'Documentation'}
(*!
<summary>No Preparation phase is needed.</summary>
*)
{endregion}
METHOD PROTECTED ProcessPreparations
VAR_INPUT
    // SA0033: Required hook; this test has no Preparation phase.
    {attribute 'analysis' := '-33'}
    Enable : BOOL; //! Phase permission supplied by the owning Test Case; FALSE does not authorize progression, while observation may continue.
END_VAR
END_METHOD

{region 'Documentation'}
(*!
<summary>Restarts the scenario sequence and outer checks.</summary>
*)
{endregion}
METHOD PROTECTED ProcessReset
FScenario := ScenarioFirstOfMultiple;
FChecked := FALSE;
FSubjectEnable := FALSE;
FContinueScenario := FALSE;
FEvaluateSubjects := FALSE;
FObservationReady := FALSE;
FFirstFailedScenario := 0;
FFailedDuringEvaluation := FALSE;
FCapture.Reset();
ResetSubjects();
FResults.Reset();
FActivity.Reset();
FInputs.Reset();
FFindings.Reset();
CompleteReset();
END_METHOD

{region 'Documentation'}
(*!
<summary>Consumes reset before each independent scenario; continuation retains subject state.</summary>
*)
{endregion}
METHOD PROTECTED ProcessTests
VAR_INPUT
    Enable : BOOL; //! Phase permission supplied by the owning Test Case; FALSE does not authorize progression, while observation may continue.
END_VAR
IF NOT Enable THEN
    RETURN;
END_IF;

IF FChecked THEN
    FChecked := FALSE;
    FObservationReady := FALSE;
    IF FEvaluateSubjects THEN
        IF FScenario = LastScenario THEN
            CompleteTests();
            RETURN;
        END_IF;
        FScenario := FScenario + 1;
    END_IF;
    FEvaluateSubjects := NOT FEvaluateSubjects;
END_IF;

IF NOT SelectScenario() THEN
    RETURN;
END_IF;
IF FContinueScenario THEN
    FEvaluateSubjects := TRUE;
END_IF;
FCapture.Reset();
IF NOT FEvaluateSubjects THEN
    ResetSubjects();
END_IF;
FDataBefore := FData;
FWideDataBefore := FWideData;
FTokenBefore := FToken;
FWideTokenBefore := FWideToken;
CallSubjects();
CheckResults();
FInputsMatch := (FData[-2] = FDataBefore[-2])
    AND (FData[-1] = FDataBefore[-1])
    AND (FData[0] = FDataBefore[0])
    AND (FData[1] = FDataBefore[1])
    AND (FData[2] = FDataBefore[2])
    AND (FData[3] = FDataBefore[3])
    AND (FWideData[-2] = FWideDataBefore[-2])
    AND (FWideData[-1] = FWideDataBefore[-1])
    AND (FWideData[0] = FWideDataBefore[0])
    AND (FWideData[1] = FWideDataBefore[1])
    AND (FWideData[2] = FWideDataBefore[2])
    AND (FWideData[3] = FWideDataBefore[3])
    AND (FToken[4] = FTokenBefore[4])
    AND (FToken[5] = FTokenBefore[5])
    AND (FWideToken[-5] = FWideTokenBefore[-5])
    AND (FWideToken[-4] = FWideTokenBefore[-4]);
CheckFindings();
IF (FFirstFailedScenario = 0)
    AND NOT (FResultsMatch AND FActivityMatch AND FInputsMatch AND FFindingsMatch) THEN
    FFirstFailedScenario := FScenario;
    FFailedDuringEvaluation := FEvaluateSubjects;
END_IF;
FObservationReady := TRUE;
END_METHOD

{region 'Documentation'}
(*!
<summary>Queues reset; the next bound FB call consumes it without evaluating.</summary>
*)
{endregion}
METHOD PRIVATE ResetSubjects
FValue.Reset();
FWideValue.Reset();
FArray.Reset();
FWideArray.Reset();
END_METHOD

{region 'Documentation'}
(*!
<summary>Selects explicit stimuli and expected results for one scenario.</summary>
*)
{endregion}
METHOD PRIVATE SelectScenario : BOOL //! TRUE after selecting a supported scenario and its literal expectations; FALSE reports an unknown scenario.
SelectScenario := FALSE;
FSubjectEnable := TRUE;
FContinueScenario := FALSE;
FData[-2] := 9;
FData[-1] := 1;
FData[0] := 2;
FData[1] := 1;
FData[2] := 2;
FData[3] := 9;
FWideData[-2] := WORD#16#0009;
FWideData[-1] := WORD#16#0101;
FWideData[0] := WORD#16#0202;
FWideData[1] := WORD#16#0101;
FWideData[2] := WORD#16#0202;
FWideData[3] := WORD#16#0009;
FToken[4] := 1;
FToken[5] := 2;
FWideToken[-5] := WORD#16#0101;
FWideToken[-4] := WORD#16#0202;
FStartIndex := -2;
FLength := 6;
FExpected := 1;
FValueToken := 1;
FWideValueToken := WORD#16#0101;
FMask := BYTE#16#FF;
FWideMask := WORD#16#FFFF;
CASE FScenario OF
    ScenarioFirstOfMultiple:
        FValueExpectedResult := E_Result.Passed;
        FValueExpectedFinding := FALSE;
        FWideValueExpectedResult := E_Result.Failed;
        FWideValueExpectedFinding := TRUE;
        FArrayExpectedResult := E_Result.Failed;
        FArrayExpectedFinding := TRUE;
        FWideArrayExpectedResult := E_Result.Passed;
        FWideArrayExpectedFinding := FALSE;
    ScenarioAtStart:
        FStartIndex := -1;
        FLength := 5;
        FExpected := 0;
        FValueExpectedResult := E_Result.Passed;
        FValueExpectedFinding := FALSE;
        FWideValueExpectedResult := E_Result.Failed;
        FWideValueExpectedFinding := TRUE;
        FArrayExpectedResult := E_Result.Failed;
        FArrayExpectedFinding := TRUE;
        FWideArrayExpectedResult := E_Result.Passed;
        FWideArrayExpectedFinding := FALSE;
    ScenarioLastCandidate:
        FStartIndex := 0;
        FLength := 3;
        FExpected := 1;
        FValueExpectedResult := E_Result.Passed;
        FValueExpectedFinding := FALSE;
        FWideValueExpectedResult := E_Result.Failed;
        FWideValueExpectedFinding := TRUE;
        FArrayExpectedResult := E_Result.Failed;
        FArrayExpectedFinding := TRUE;
        FWideArrayExpectedResult := E_Result.Passed;
        FWideArrayExpectedFinding := FALSE;
    ScenarioDistanceMismatch:
        FExpected := 2;
        FValueExpectedResult := E_Result.Failed;
        FValueExpectedFinding := TRUE;
        FWideValueExpectedResult := E_Result.Passed;
        FWideValueExpectedFinding := FALSE;
        FArrayExpectedResult := E_Result.Passed;
        FArrayExpectedFinding := FALSE;
        FWideArrayExpectedResult := E_Result.Failed;
        FWideArrayExpectedFinding := TRUE;
    ScenarioElementDistance:
        FData[-1] := 9;
        FData[0] := 9;
        FWideData[-1] := 9;
        FWideData[0] := 9;
        FExpected := 3;
        FValueExpectedResult := E_Result.Passed;
        FValueExpectedFinding := FALSE;
        FWideValueExpectedResult := E_Result.Failed;
        FWideValueExpectedFinding := TRUE;
        FArrayExpectedResult := E_Result.Failed;
        FArrayExpectedFinding := TRUE;
        FWideArrayExpectedResult := E_Result.Passed;
        FWideArrayExpectedFinding := FALSE;
    ScenarioMaskedValue:
        FData[-2] := BYTE#16#81;
        FWideData[-2] := WORD#16#8001;
        FMask := BYTE#16#0F;
        FWideMask := WORD#16#000F;
        FExpected := 0;
        FValueExpectedResult := E_Result.Passed;
        FValueExpectedFinding := FALSE;
        FWideValueExpectedResult := E_Result.Failed;
        FWideValueExpectedFinding := TRUE;
        FArrayExpectedResult := E_Result.Passed;
        FArrayExpectedFinding := FALSE;
        FWideArrayExpectedResult := E_Result.Failed;
        FWideArrayExpectedFinding := TRUE;
    ScenarioLastValue:
        FStartIndex := 0;
        FLength := 4;
        FValueToken := 9;
        FWideValueToken := 9;
        FExpected := 3;
        FValueExpectedResult := E_Result.Passed;
        FValueExpectedFinding := FALSE;
        FWideValueExpectedResult := E_Result.Failed;
        FWideValueExpectedFinding := TRUE;
        FArrayExpectedResult := E_Result.Passed;
        FArrayExpectedFinding := FALSE;
        FWideArrayExpectedResult := E_Result.Failed;
        FWideArrayExpectedFinding := TRUE;
    ScenarioAbsent:
        FValueToken := 7;
        FWideValueToken := 7;
        FToken[4] := 7;
        FWideToken[-5] := 7;
        FValueExpectedResult := E_Result.Failed;
        FValueExpectedFinding := TRUE;
        FWideValueExpectedResult := E_Result.Failed;
        FWideValueExpectedFinding := TRUE;
        FArrayExpectedResult := E_Result.Failed;
        FArrayExpectedFinding := TRUE;
        FWideArrayExpectedResult := E_Result.Failed;
        FWideArrayExpectedFinding := TRUE;
    ScenarioTokenTooLong:
        FLength := 1;
        FValueToken := 9;
        FWideValueToken := 9;
        FExpected := 0;
        FValueExpectedResult := E_Result.Passed;
        FValueExpectedFinding := FALSE;
        FWideValueExpectedResult := E_Result.Failed;
        FWideValueExpectedFinding := TRUE;
        FArrayExpectedResult := E_Result.Error;
        FArrayExpectedFinding := TRUE;
        FWideArrayExpectedResult := E_Result.Error;
        FWideArrayExpectedFinding := TRUE;
    ScenarioEmptyRange:
        FLength := 0;
        FValueExpectedResult := E_Result.Error;
        FValueExpectedFinding := TRUE;
        FWideValueExpectedResult := E_Result.Error;
        FWideValueExpectedFinding := TRUE;
        FArrayExpectedResult := E_Result.Error;
        FArrayExpectedFinding := TRUE;
        FWideArrayExpectedResult := E_Result.Error;
        FWideArrayExpectedFinding := TRUE;
    ScenarioRangePastEnd:
        FStartIndex := 3;
        FLength := 2;
        FValueExpectedResult := E_Result.Error;
        FValueExpectedFinding := TRUE;
        FWideValueExpectedResult := E_Result.Error;
        FWideValueExpectedFinding := TRUE;
        FArrayExpectedResult := E_Result.Error;
        FArrayExpectedFinding := TRUE;
        FWideArrayExpectedResult := E_Result.Error;
        FWideArrayExpectedFinding := TRUE;
ELSE
    Error(Message := 'Unknown Assertion scenario.');
    RETURN;
END_CASE;
SelectScenario := TRUE;
END_METHOD

END_FUNCTION_BLOCK

// ---- SelfTests/TestSuites/TestSuite_AssertionArrays.TcPOU
{region 'Documentation'}
(*!
<summary>Checks array comparison and search boundaries with isolated Assertion subjects.</summary>
*)
{endregion}
FUNCTION_BLOCK TestSuite_AssertionArrays EXTENDS TestSuiteBase
VAR
    FArrayComparison : Test_AssertionArrayComparison;
    FArrayValueSearch : Test_AssertionArrayValueSearch;
    FArrayPatternSearch : Test_AssertionArrayPatternSearch;
    FMaskedArrayComparison : Test_AssertionMaskedArrayComparison;
    FFloatingPointArray : Test_AssertionFloatingPointArray;
    FArrayTextBridge : Test_AssertionArrayTextBridge;
    FTestCases : ARRAY[1..TestCaseCapacity] OF I_TestCase;
END_VAR
VAR CONSTANT
    TestCaseCapacity : UINT := 6;
END_VAR

SUPER^();

{region 'Documentation'}
(*!
<summary>Initializes six isolated array comparison and search Test Cases and registers them serially.</summary>
*)
{endregion}
METHOD PROTECTED Configure
VAR_IN_OUT
    // SA0167: Borrowed owner builder; no temporary instance is created.
    {attribute 'analysis' := '-167'}
    Builder : TestSuiteConfigurationBuilder; //! Borrowed owner configuration builder used only during this Configure call; register this owner's concrete children.
END_VAR
VAR
    TestConfig : ST_TestCaseConfig;
END_VAR
Builder.Initialize(Mode := E_OrchestrationMode.Serial,
    TestCases := FTestCases);
FArrayComparison.Initialize(Parent := THIS^,
    TestName := 'ArrayComparison',
    Config := TestConfig);
Builder.Register(TestCase := FArrayComparison);
FArrayValueSearch.Initialize(Parent := THIS^,
    TestName := 'ArrayValueSearch',
    Config := TestConfig);
Builder.Register(TestCase := FArrayValueSearch);
FArrayPatternSearch.Initialize(Parent := THIS^,
    TestName := 'ArrayPatternSearch',
    Config := TestConfig);
Builder.Register(TestCase := FArrayPatternSearch);
FMaskedArrayComparison.Initialize(Parent := THIS^,
    TestName := 'MaskedArrayComparison',
    Config := TestConfig);
Builder.Register(TestCase := FMaskedArrayComparison);
FFloatingPointArray.Initialize(Parent := THIS^,
    TestName := 'FloatingPointArray',
    Config := TestConfig);
Builder.Register(TestCase := FFloatingPointArray);
FArrayTextBridge.Initialize(Parent := THIS^,
    TestName := 'ArrayTextBridge',
    Config := TestConfig);
Builder.Register(TestCase := FArrayTextBridge);
END_METHOD

{region 'Documentation'}
(*!
<summary>Returns a registered scenario using its original array index.</summary>
*)
{endregion}
METHOD PUBLIC GetTestCase : I_TestCase //! Typed child interface at the original array index; zero when no entry is available.
VAR_INPUT
    Index : DINT; //! Original occupied child-array index, rather than an ordinal position.
END_VAR
GetTestCase := 0;
IF (ChildCount = 0) OR (Index < ChildArrayLowerBound)
    OR (DINT_TO_LINT(Index) >= DINT_TO_LINT(ChildArrayLowerBound) + UINT_TO_LINT(ChildCount)) THEN
    RETURN;
END_IF;
GetTestCase := FTestCases[Index];
END_METHOD

{region 'Documentation'}
(*!
<summary>Calls every owned scenario once per initialized Suite cycle.</summary>
*)
{endregion}
METHOD PROTECTED ProcessTestCases
FArrayComparison();
FArrayValueSearch();
FArrayPatternSearch();
FMaskedArrayComparison();
FFloatingPointArray();
FArrayTextBridge();
END_METHOD

END_FUNCTION_BLOCK

// ---- SelfTests/TestCases/TestSuite_AssertionArrays/Test_AssertionArrayComparison.TcPOU
{region 'Documentation'}
(*!
<summary>Checks selected-region INT equality and BOOL all-elements equality.</summary>
<description>
Independent scenarios use a bound reset call followed by an evaluation call.
ProcessAssertions checks each observation before ProcessTests advances.
SelectScenario defines literal expected results; production algorithms are inherited.
Only the explicitly marked continuation retains a previous subject result.
Inputs belong to this Test Case and are compared with their pre-call values.
Expected subject findings remain in the local capture, never the outer event stream.
FirstFailedScenario and FailedDuringEvaluation retain the first mismatch.
</description>
*)
{endregion}
FUNCTION_BLOCK Test_AssertionArrayComparison EXTENDS TestCaseBase
VAR
    FEqual : AssertEqualArray_Int;
    FEqualExpectedResult : E_Result;
    FEqualExpectedFinding : BOOL;
    FAll : AssertArrayAllEqual_Bool;
    FAllExpectedResult : E_Result;
    FAllExpectedFinding : BOOL;
    FData : ARRAY[-3..3] OF INT;
    FDataBefore : ARRAY[-3..3] OF INT;
    FExpected : ARRAY[5..7] OF INT;
    FExpectedBefore : ARRAY[5..7] OF INT;
    FSingleExpected : ARRAY[9..9] OF INT;
    FSingleExpectedBefore : ARRAY[9..9] OF INT;
    FFlags : ARRAY[-1..2] OF BOOL;
    FFlagsBefore : ARRAY[-1..2] OF BOOL;
    FStartIndex : DINT;
    FBoolStartIndex : DINT;
    FLength : USINT;
    FUseSingleExpected : BOOL;
    FSubjectEnable : BOOL;
    FContinueScenario : BOOL;
    FCapture : EventBuffer;
    FEvents : ARRAY[1..CaptureLength] OF ST_Event;
    FCaptureFifo : ST_FifoStatus;
    FCaptureStatus : ST_EventBufferStatus;
    FSetupValid : BOOL;
    FScenario : UINT;
    FChecked : BOOL;
    FEvaluateSubjects : BOOL;
    FObservationReady : BOOL;
    FFirstFailedScenario : UINT;
    FFailedDuringEvaluation : BOOL;
    FResultsMatch : BOOL;
    FResults : AssertTrue;
    FActivityMatch : BOOL;
    FActivity : AssertTrue;
    FInputsMatch : BOOL;
    FInputs : AssertTrue;
    FFindingsMatch : BOOL;
    FFindings : AssertTrue;
END_VAR
VAR CONSTANT
    CaptureLength : UINT := 8;
    ScenarioSelectedRegion : UINT := 1;
    ScenarioFirstMismatch : UINT := 2;
    ScenarioLastMismatch : UINT := 3;
    ScenarioLowerBoundary : UINT := 4;
    ScenarioUpperBoundary : UINT := 5;
    ScenarioSingleElement : UINT := 6;
    ScenarioBelowLowerBound : UINT := 7;
    ScenarioAboveUpperBound : UINT := 8;
    ScenarioEndOutsideRange : UINT := 9;
    ScenarioEmptyRange : UINT := 10;
    ScenarioMismatchBeforeInvalidRange : UINT := 11;
    ScenarioInvalidRangeAfterFailure : UINT := 12;
    LastScenario : UINT := ScenarioInvalidRangeAfterFailure;
END_VAR

SUPER^();

{region 'Documentation'}
(*!
<summary>Aggregates only outer checks, not intentionally failing subjects.</summary>
*)
{endregion}
METHOD PROTECTED AggregateResults
VAR_INPUT
    Aggregator : I_ResultAggregator; //! Borrowed result sink owned by the outer Test Case; add this test's checking Assertions without resetting or retaining the sink.
END_VAR
Aggregator.AddProvider(Provider := FResults);
Aggregator.AddProvider(Provider := FActivity);
Aggregator.AddProvider(Provider := FInputs);
Aggregator.AddProvider(Provider := FFindings);
END_METHOD

{region 'Documentation'}
(*!
<summary>Calls each inherited production subject once with caller-owned input storage.</summary>
*)
{endregion}
METHOD PRIVATE CallSubjects
IF FUseSingleExpected THEN
    FEqual(Enable := FSubjectEnable,
        State := E_State.Running,
        StartIndex := FStartIndex,
        IN := FData,
        Expected := FSingleExpected);
ELSE
    FEqual(Enable := FSubjectEnable,
        State := E_State.Running,
        StartIndex := FStartIndex,
        IN := FData,
        Expected := FExpected);
END_IF;
FAll(Enable := FSubjectEnable,
    State := E_State.Running,
    StartIndex := FBoolStartIndex,
    Length := FLength,
    Expected := TRUE,
    IN := FFlags);
END_METHOD

{region 'Documentation'}
(*!
<summary>Checks one subject finding in call order; expected outcomes come from the scenario.</summary>
*)
{endregion}
METHOD PRIVATE CheckFinding : BOOL //! TRUE when the required finding checks pass; calls requiring no finding also succeed.
VAR_INPUT
    Subject : I_Assertion; //! Assertion interface supplying the expected finding identity.
    ExpectedResult : E_Result; //! Independently authored result expected in the captured finding.
    ExpectedFinding : BOOL; //! TRUE when this scenario requires a finding during active evaluation.
END_VAR
VAR_IN_OUT
    Index : UINT; //! One-based next finding index; advanced when this call checks a required finding.
END_VAR
CheckFinding := TRUE;
IF FEvaluateSubjects AND ExpectedFinding THEN
    CheckFinding := (FEvents[Index].SequenceId = UINT_TO_UDINT(Index))
        AND (FEvents[Index].Name = Subject.Name)
        AND (FEvents[Index].OwnerScope = E_OwnerScope.Assertion)
        AND (FEvents[Index].EventType = E_EventType.Result)
        AND (FEvents[Index].State = E_State.Running)
        AND (FEvents[Index].Result = ExpectedResult)
        AND (FEvents[Index].Message <> '');
    Index := Index + 1;
END_IF;
END_METHOD

